//---------------------------------------------------------VFD
    // VTD (MOVI-C MOVIPRO) / Module 1 (Standard 8 PD), MOVIKIT Positioning Drive.
    // Raw 16-bit UINT data, as defined in SpaceX.tsproj; no scaling or decoding.
    // Link each variable to the channel with the same number in TwinCAT XAE.
    // Word meanings from MOVISUITE; bit meanings and units still pending SEW.

    // Drive -> PLC: Inputs 8 PD / PDO 16#1A02 / object 16#7002.
    // Read only by FC Inputs, into Control.VTD.Motor.stProcessInput.
    VTD_PI_01 AT %I* : UINT; // PI 1, 16#7002:01 - Status word
    VTD_PI_02 AT %I* : UINT; // PI 2, 16#7002:02 - Actual speed
    VTD_PI_03 AT %I* : UINT; // PI 3, 16#7002:03 - Status/main fault - subfault
    VTD_PI_04 AT %I* : UINT; // PI 4, 16#7002:04 - Torque
    VTD_PI_05 AT %I* : UINT; // PI 5, 16#7002:05 - Digital inputs
    VTD_PI_06 AT %I* : UINT; // PI 6, 16#7002:06 - Actual application mode
    VTD_PI_07 AT %I* : UINT; // PI 7, 16#7002:07 - Actual position high word (DL50)
    VTD_PI_08 AT %I* : UINT; // PI 8, 16#7002:08 - Actual position low word (DL50)

    // PLC -> drive: Outputs 8 PD / PDO 16#1602 / object 16#6002.
    // Written only by FC Outputs, from Control.VTD.Motor.aProcessOutput.
    VTD_PO_01 AT %Q* : UINT; // PO 1, 16#6002:01 - Control word
    VTD_PO_02 AT %Q* : UINT; // PO 2, 16#6002:02 - Setpoint speed
    VTD_PO_03 AT %Q* : UINT; // PO 3, 16#6002:03 - Setpoint acceleration
    VTD_PO_04 AT %Q* : UINT; // PO 4, 16#6002:04 - Setpoint deceleration
    VTD_PO_05 AT %Q* : UINT; // PO 5, 16#6002:05 - Digital outputs
    VTD_PO_06 AT %Q* : UINT; // PO 6, 16#6002:06 - Setpoint application mode
    VTD_PO_07 AT %Q* : UINT; // PO 7, 16#6002:07 - Target position high word
    VTD_PO_08 AT %Q* : UINT; // PO 8, 16#6002:08 - Target position low word

    // EtherCAT diagnostics of the VTD box. Not linked yet: link manually in XAE.
    // Read only by FC Inputs.
    VTD_WcState AT %I* : BOOL; // VTD > WcState > WcState (TRUE = data invalid)
    VTD_EcState AT %I* : UINT; // VTD > InfoData > State (8 = OP)
	
	//----------------------------------------------------EXTRACTOR CONVEYOR
END_VAR

// ---- GVLs/Settings.TcGVL
{attribute 'qualified_only'}
VAR_GLOBAL
	VTD:  VTD_Settings_DUT;
	ECnv:  ECnv_Settings_DUT;
	LCnv:  ARRAY[1..6] OF Buffer_Cnv_Settings_DUT;
	Turn_Table: Turn_Table_Settings_DUT;
	TBCnv:  TBCnv_Settings_DUT;
	Pop_Up_Cnv: ARRAY[1..2] OF PopUp_Settings_DUT;
	Roller_Cnv: ARRAY[1..5] OF Roller_Settings_DUT;
	Chain_Cnv: Chain_Settings_DUT;
// 	Shuttle_MQTT:  MQTT_Settings;
	System:  System_Settings_DUT;
END_VAR

// ---- GVLs/System.TcGVL
{attribute 'qualified_only'}
VAR_GLOBAL
	Id:  UINT;
	CancelOrders:  BOOL;
	PauseOrders:  Bool;
	ResumeOrders:  Bool;
	OrderSent:  Bool;
	CurrentOrder:  UInt;
	NextOrder:  UInt;
	OrderTable:  ARRAY[0..99] OF OrderTable_DUT;
	StepTable:  ARRAY[0..20] OF OrderTable_DUT;
	CarParked_Confirm:  Bool;
	Running:  Bool;
	IDLE:  Bool;
	Error:  Bool;
	State:  USInt;
	ResetError:  Bool;
	Ready:  Bool;
	Selected:  Bool;
	Auto_Man:  Bool;
	Paused:  Bool;
// 	Watchdog_TimeOut:  STRUCT;
END_VAR

// ---- GVLs/System_Control.TcGVL
{attribute 'qualified_only'}
VAR_GLOBAL
	Reset_All:  BOOL;
	MQTT_Enable:  BOOL;
	OPC_Enable:  Bool;
END_VAR

// ---- POUs/MAIN.TcPOU
PROGRAM MAIN
VAR
	 // TEST ONLY - VTD MOVIPRO process data communication check.
    fbVtdProcessDataTest : FB_SEW_ProcessDataTest;
    // TEST ONLY - VTD manual control from the screen VTD_ManualTest.
    fbVtdManualControl : FB_VTD_ManualControl;
    // Safety reset from the HMI (button SAFETY RESET): one pulse per rising edge.
    rtSafetyReset : R_TRIG;
    tpSafetyReset : TP;
END_VAR

run := TRUE;

// 1. IO inputs -> internal variables
Inputs();

// 2. Logic on internal variables
// Safety reset from the HMI: one 500 ms pulse on IO_Safety.ErrorAcknowledgement and
// IO_Safety.SEW_Safety_Reset (written in Outputs). It is a request only: the TwinSAFE
// logic accepts it or not. Holding the button does not repeat the reset.
rtSafetyReset(CLK := GVL_HMI_System.stCommand.bSafetyReset);
tpSafetyReset(IN := rtSafetyReset.Q, PT := T#500MS);
Control.SafetyReset := tpSafetyReset.Q;

// TEST ONLY - two sources can write the VTD process outputs, only one at a time:
//  - the raw write of the process data screen is refused (its HMI toggle is reset)
//    while the manual screen has the drive enabled;
//  - the manual control is inhibited while the raw write is active.
IF fbVtdManualControl.q_stStatus.bEnableActive THEN
    GVL_HMI_VTD.stPdCommand.bTestWriteEnable := FALSE;
END_IF

// TEST ONLY - VTD MOVIPRO process data communication check.
fbVtdProcessDataTest(
    i_aProcessInput := Control.VTD.Motor.stProcessInput.aWord,
    i_bWcStateError := Control.VTD.Motor.stProcessInput.bWcStateError,
    i_uiEcState := Control.VTD.Motor.stProcessInput.uiEcState,
    i_bTestWriteEnable := GVL_HMI_VTD.stPdCommand.bTestWriteEnable,
    i_bTestAllowControlWord := GVL_HMI_VTD.stPdCommand.bTestAllowControlWord,
    i_aTestProcessOutput := GVL_HMI_VTD.stPdCommand.aTestProcessOutput);

// TEST ONLY - VTD manual control (jog, modes, speed, software stop, reset).
fbVtdManualControl(
    i_stProcessInput := Control.VTD.Motor.stProcessInput,
    i_bInhibit := fbVtdProcessDataTest.q_bTestWriteActive,
    i_stSettings := GVL_HMI_VTD.stManualSettings,
    io_stCommand := GVL_HMI_VTD.stManualCommand);

IF fbVtdProcessDataTest.q_bTestWriteActive THEN
    Control.VTD.Motor.aProcessOutput := fbVtdProcessDataTest.q_aProcessOutput;
ELSE
    Control.VTD.Motor.aProcessOutput := fbVtdManualControl.q_aProcessOutput;
END_IF

// 3. HMI status
FC_VTD_PdHmiUpdateStatus(
    io_fbProcessData := fbVtdProcessDataTest,
    io_stStatus := GVL_HMI_VTD.stPdStatus);
// PO really sent to the drive (raw write or manual control).
GVL_HMI_VTD.stPdStatus.aProcessOutputSent := Control.VTD.Motor.aProcessOutput;
GVL_HMI_VTD.stManualStatus := fbVtdManualControl.q_stStatus;
GVL_HMI_System.stStatus.bSafetyResetActive := tpSafetyReset.Q;

// 4. Internal variables -> IO outputs
Outputs();

END_PROGRAM

// ---- POUs/SEW/FB_SEW_ProcessDataTest.TcPOU
// TEST ONLY - communication check between TwinCAT and a MOVIPRO running
// MOVIKIT Positioning Drive with the "Standard 8 PD" fieldbus interface.
//
// PD layout confirmed from MOVISUITE (VTD > MOVIKIT Positioning Drive > Basic settings):
//   PO 1 Control word              PI 1 Status word
//   PO 2 Setpoint speed            PI 2 Actual speed
//   PO 3 Setpoint acceleration     PI 3 Status/main fault - subfault
//   PO 4 Setpoint deceleration     PI 4 Torque (selectable in MOVISUITE)
//   PO 5 Digital outputs           PI 5 Digital inputs
//   PO 6 Setpoint application mode PI 6 Actual application mode
//   PO 7 Target position high word PI 7 Actual position high word
//   PO 8 Target position low word  PI 8 Actual position low word
//
// NOT yet confirmed (pending SEW): control/status word bit meanings,
// application mode values, user units and scaling of speed, ramps, torque and
// position. All decoded values are therefore RAW and carry no engineering unit.
//
// This block does not control the drive. All process outputs are 0 unless a
// TEST ONLY write is explicitly enabled online. The control word (PO 1) stays 0
// unless it is separately enabled. A control word of 0 is not confirmed as a
// safe state for this vertical axis; confirm with SEW before writing anything.
FUNCTION_BLOCK FB_SEW_ProcessDataTest
VAR_INPUT
    i_aProcessInput : ARRAY[1..8] OF UINT;      // PI 1..8, raw from the drive
    i_bWcStateError : BOOL;                     // EtherCAT WcState of the drive box (TRUE = data invalid)
    i_uiEcState : UINT;                         // EtherCAT InfoData.State of the drive box (8 = OP)

    i_bTestWriteEnable : BOOL;                  // TEST ONLY - allow PO 2..8 to be written
    i_bTestAllowControlWord : BOOL;             // TEST ONLY - additionally allow PO 1 (control word)
    i_aTestProcessOutput : ARRAY[1..8] OF UINT; // TEST ONLY - raw values to send to PO 1..8
    i_tTestWriteTimeout : TIME := T#10M;        // TEST ONLY write is dropped after this time
END_VAR
VAR_OUTPUT
    q_bCommunicationOk : BOOL;                  // Drive in OP and working counter valid
    q_udiInputChangeCount : UDINT;              // Cycles in which any PI word changed (wraps)

    q_wStatusWord : WORD;                       // PI 1, bit meanings pending SEW
    q_iActualSpeedRaw : INT;                    // PI 2, signed assumed, unit pending SEW
    q_wFaultCode : WORD;                        // PI 3, main fault / subfault, raw
    q_iTorqueRaw : INT;                         // PI 4, signed assumed, unit pending SEW
    q_wDigitalInputs : WORD;                    // PI 5, raw
    q_uiActualApplicationMode : UINT;           // PI 6, value meanings pending SEW
    q_diActualPositionRaw : DINT;               // PI 7 (high) + PI 8 (low), user units pending SEW

    q_bTestWriteActive : BOOL;                  // TEST ONLY write currently applied
    q_bTestWriteExpired : BOOL;                 // Timeout elapsed; toggle i_bTestWriteEnable to restart
    q_tTestWriteElapsed : TIME;                 // Elapsed time of the current TEST ONLY write window
    q_aProcessOutput : ARRAY[1..8] OF UINT;     // PO 1..8, raw to the drive
END_VAR
VAR
    aPreviousInput : ARRAY[1..8] OF UINT;
    bInputChanged : BOOL;
    dwActualPosition : DWORD;
    iWord : INT;

    rtrigTestWriteEnable : R_TRIG;
    tonTestWriteTimeout : TON;
END_VAR

// Communication status: EtherCAT state OP (lower nibble = 8) and valid working counter.
q_bCommunicationOk := (NOT i_bWcStateError) AND ((i_uiEcState AND 16#000F) = 8);

// Count cycles in which the drive sends new data. A counter that keeps rising
// while the drive is powered shows that PI data really arrives.
bInputChanged := FALSE;
FOR iWord := 1 TO 8 DO
    IF i_aProcessInput[iWord] <> aPreviousInput[iWord] THEN
        bInputChanged := TRUE;
    END_IF
END_FOR
aPreviousInput := i_aProcessInput;

IF bInputChanged THEN
    q_udiInputChangeCount := q_udiInputChangeCount + 1;
END_IF

// Raw decoding. Same-size integer conversions keep the bit pattern.
q_wStatusWord := UINT_TO_WORD(i_aProcessInput[1]);
q_iActualSpeedRaw := UINT_TO_INT(i_aProcessInput[2]);
q_wFaultCode := UINT_TO_WORD(i_aProcessInput[3]);
q_iTorqueRaw := UINT_TO_INT(i_aProcessInput[4]);
q_wDigitalInputs := UINT_TO_WORD(i_aProcessInput[5]);
q_uiActualApplicationMode := i_aProcessInput[6];

// Position word order (PI 7 = high, PI 8 = low) is shown in MOVISUITE.
// Signed 32-bit integer: numeric value, not an IEEE-754 bit pattern.
dwActualPosition := SHL(UINT_TO_DWORD(i_aProcessInput[7]), 16)
                    OR UINT_TO_DWORD(i_aProcessInput[8]);
q_diActualPositionRaw := DWORD_TO_DINT(dwActualPosition);

// TEST ONLY write enable with timeout. A rising edge restarts the timeout.
rtrigTestWriteEnable(CLK := i_bTestWriteEnable);
IF rtrigTestWriteEnable.Q THEN
    q_bTestWriteExpired := FALSE;
END_IF

tonTestWriteTimeout(IN := i_bTestWriteEnable AND NOT q_bTestWriteExpired,
                    PT := i_tTestWriteTimeout);
IF tonTestWriteTimeout.Q THEN
    q_bTestWriteExpired := TRUE;
END_IF
q_tTestWriteElapsed := tonTestWriteTimeout.ET;

q_bTestWriteActive := i_bTestWriteEnable AND NOT q_bTestWriteExpired;

// Process outputs: 0 by default.
FOR iWord := 1 TO 8 DO
    q_aProcessOutput[iWord] := 0;
END_FOR

IF q_bTestWriteActive THEN
    FOR iWord := 2 TO 8 DO
        q_aProcessOutput[iWord] := i_aTestProcessOutput[iWord];
    END_FOR

    IF i_bTestAllowControlWord THEN
        q_aProcessOutput[1] := i_aTestProcessOutput[1];
    END_IF
END_IF

END_FUNCTION_BLOCK

// ---- POUs/VTD/FB_VTD_ManualControl.TcPOU
// TEST ONLY - manual control of the VTD MOVIPRO from the screen VTD_ManualTest.
// Temporary owner of the axis for commissioning; VTD_FB replaces it in production.
// Uses FB_SEW_Drive (MOVIKIT Positioning Drive, Standard 8 PD, SEW manual 33959862).
//
// Behavior:
//  - ENABLE is a request from the HMI. It is dropped, and the HMI toggle reset, on
//    software stop, communication loss, drive error, STO active or while the raw
//    process data write is active. No automatic restart.
//    ENABLE off while turning: stop with the PO 4 ramp first, then remove the enable.
//  - JOG -/+ (modes 100/101) is hold-to-run. A button must be released before it is
//    accepted, and it is ignored after tJogMaxTime until it is released.
//  - RUN -/+ (mode 200) and START (modes 300/400/401) are latched; STOP clears them
//    (deceleration with PO 4). Reversing in mode 200 requires STOP first.
//  - The target position is taken from the HMI only with START.
//  - The operating mode changes only at standstill without motion command,
//    because the drive stops when PO 6 changes (manual chapter 8.1).
//  - Speed = iSpeedPercent (0..100 %) of stManualSettings.iMaxSpeed (user units).
//  - SOFTWARE STOP is NOT an emergency stop and not a safety function. It removes the
//    enable, so the drive stops with FCB 14 (emergency stop ramp) and applies the brake.
//    The safety-rated stop is the hardwired / TwinSAFE emergency stop (STO).
//  - RESET clears the software stop and sends a drive fault reset pulse (PO 1.8).
//  - Never used: release brake without enable, output stage inhibit, deactivation of
//    the software limit switches (not set by FB_SEW_Drive).
//
// Drive status is evaluated from the previous call of FB_SEW_Drive (one PLC cycle).
FUNCTION_BLOCK FB_VTD_ManualControl
VAR_INPUT
    i_stProcessInput : ST_SEW_ProcessInput8;  // Raw PI 1..8 + EtherCAT diagnostics (Control.VTD.Motor)
    i_bInhibit : BOOL;                        // TRUE = another source writes the PO (raw PD test); enable is dropped
    i_stSettings : ST_VTD_ManualSettings;     // Max speed, ramps (user units) and jog max time
END_VAR
VAR_IN_OUT
    io_stCommand : ST_VTD_ManualHmiCommand;   // HMI commands; bEnable, eModeRequest and iSpeedPercent are written back
END_VAR
VAR_OUTPUT
    q_aProcessOutput : ARRAY[1..8] OF UINT;   // Raw PO 1..8 (to Control.VTD.Motor.aProcessOutput)
    q_stStatus : ST_VTD_ManualHmiStatus;      // To GVL_HMI_VTD.stManualStatus
END_VAR
VAR
    fbDrive : FB_SEW_Drive;
    eModeActive : E_SEW_MovikitMode := E_SEW_MovikitMode.JogSpeedControlled;

    // Operating mode
    bModeSupported : BOOL;
    bModeChangeAllowed : BOOL;
    bModeRejected : BOOL;
    bJogMode : BOOL;
    bSpeedMode : BOOL;
    bReferencingMode : BOOL;
    bPositioningMode : BOOL;

    // Enable
    bSoftwareStopLatched : BOOL;
    bSettingsValid : BOOL;
    bEnableBlocked : BOOL;
    bEnableRequest : BOOL;
    bEnableActive : BOOL;

    // Motion commands
    bMotionCommand : BOOL;
    bJogButtonsReleased : BOOL;
    bJogArmed : BOOL;
    bJogTimeout : BOOL;
    bJogPositive : BOOL;
    bJogNegative : BOOL;
    bRunAvailable : BOOL;
    bRunPositive : BOOL;
    bRunNegative : BOOL;
    bStartAvailable : BOOL;
    bStartLatched : BOOL;
    bRelativeMoveOpen : BOOL;                 // Mode 401: distance applied, target not reached yet
    bApplyRelativeRequest : BOOL;             // Mode 401: PO 1.6 pulse starts in the next cycle
    diTargetPosition : DINT;                  // PO 7/8, user units
    diSpeedTemp : DINT;
    iSpeedMagnitude : INT;
    iSpeedSetpoint : INT;

    rtrigSoftwareStop : R_TRIG;
    rtrigReset : R_TRIG;
    rtrigRunPositive : R_TRIG;
    rtrigRunNegative : R_TRIG;
    rtrigStart : R_TRIG;
    rtrigStop : R_TRIG;
    tpFaultReset : TP;
    tpApplyRelative : TP;
    tpModeRejected : TP;
    tonJogMaxTime : TON;
    tonDisableStop : TON;
    tonRelativeDone : TON;
    tonReferencingDone : TON;
END_VAR
VAR CONSTANT
    FAULT_RESET_PULSE : TIME := T#500MS;      // PO 1.8 high time (the drive resets on the rising edge)
    APPLY_RELATIVE_PULSE : TIME := T#200MS;   // PO 1.6 high time (mode 401)
    MODE_REJECTED_MESSAGE : TIME := T#3S;     // Display time of the "mode change refused" message
    DISABLE_STOP_TIMEOUT : TIME := T#5S;      // Max time to stop with PO 4 before the enable is removed
    RELATIVE_DONE_DELAY : TIME := T#500MS;    // In position + standstill for this time = relative move done
    REFERENCING_DONE_DELAY : TIME := T#1S;    // Referenced + standstill for this time = START released
END_VAR

{region "Edge detection of the HMI buttons"}
rtrigSoftwareStop(CLK := io_stCommand.bSoftwareStop);
rtrigReset(CLK := io_stCommand.bReset);
rtrigRunPositive(CLK := io_stCommand.bRunPositive);
rtrigRunNegative(CLK := io_stCommand.bRunNegative);
rtrigStart(CLK := io_stCommand.bStart);
rtrigStop(CLK := io_stCommand.bStop);
{endregion}

{region "Software stop and reset"}
// SOFTWARE STOP is not a safety function. It removes the enable, so the drive
// stops with FCB 14 (emergency stop ramp) and applies the brake.
IF rtrigSoftwareStop.Q THEN
    bSoftwareStopLatched := TRUE;
END_IF

// RESET clears the software stop and resets drive faults with a PO 1.8 pulse.
// The enable stays off until ENABLE is pressed again.
IF rtrigReset.Q AND NOT io_stCommand.bSoftwareStop THEN
    bSoftwareStopLatched := FALSE;
END_IF
tpFaultReset(IN := rtrigReset.Q, PT := FAULT_RESET_PULSE);
{endregion}

{region "Settings"}
bSettingsValid := (i_stSettings.iMaxSpeed > 0)
                  AND (i_stSettings.uiAcceleration > 0)
                  AND (i_stSettings.uiDeceleration > 0)
                  AND (i_stSettings.tJogMaxTime > T#0S);
{endregion}

{region "Operating mode (PO 6)"}
// The drive stops when PO 6 changes (manual chapter 8.1), so the mode is changed
// only at standstill and without an active motion command.
bMotionCommand := bRunPositive OR bRunNegative OR bStartLatched
                  OR io_stCommand.bJogPositive OR io_stCommand.bJogNegative;
bModeChangeAllowed := NOT bMotionCommand AND NOT fbDrive.q_stStatus.bMotorTurning;
bModeRejected := FALSE;

IF io_stCommand.eModeRequest <> eModeActive THEN
    CASE io_stCommand.eModeRequest OF
        E_SEW_MovikitMode.JogPositionControlled,
        E_SEW_MovikitMode.JogSpeedControlled,
        E_SEW_MovikitMode.Speed,
        E_SEW_MovikitMode.ReferencingOffsetConfigured,
        E_SEW_MovikitMode.PositioningAbsolute,
        E_SEW_MovikitMode.PositioningRelative:
            bModeSupported := TRUE;
    ELSE
        bModeSupported := FALSE;
    END_CASE

    IF bModeSupported AND bModeChangeAllowed THEN
        eModeActive := io_stCommand.eModeRequest;
        bRelativeMoveOpen := FALSE;
        diTargetPosition := 0;
    ELSE
        bModeRejected := TRUE;
    END_IF
END_IF

// The HMI always shows the mode really sent to the drive.
io_stCommand.eModeRequest := eModeActive;

bJogMode := (eModeActive = E_SEW_MovikitMode.JogPositionControlled)
            OR (eModeActive = E_SEW_MovikitMode.JogSpeedControlled);
bSpeedMode := (eModeActive = E_SEW_MovikitMode.Speed);
bReferencingMode := (eModeActive = E_SEW_MovikitMode.ReferencingOffsetConfigured);
bPositioningMode := (eModeActive = E_SEW_MovikitMode.PositioningAbsolute)
                    OR (eModeActive = E_SEW_MovikitMode.PositioningRelative);
{endregion}

{region "Enable (PO 1.0 + PO 1.1)"}
// The enable request is dropped - and the HMI toggle reset - when the drive cannot
// or must not run. No automatic restart: ENABLE must be pressed again.
bEnableBlocked := bSoftwareStopLatched
                  OR i_bInhibit
                  OR NOT fbDrive.q_stStatus.bCommunicationOk
                  OR fbDrive.q_stStatus.bError
                  OR NOT fbDrive.q_stStatus.bStoInactive;

IF bEnableBlocked THEN
    io_stCommand.bEnable := FALSE;
END_IF
bEnableRequest := io_stCommand.bEnable AND NOT bEnableBlocked;

// ENABLE switched off while turning: the motion commands are cleared below, the
// drive stops with the PO 4 ramp and the enable is removed at standstill
// (at the latest after DISABLE_STOP_TIMEOUT, then FCB 14).
tonDisableStop(IN := bEnableActive AND NOT bEnableRequest AND NOT bEnableBlocked,
               PT := DISABLE_STOP_TIMEOUT);
bEnableActive := bEnableRequest
                 OR (bEnableActive
                     AND NOT bEnableBlocked
                     AND fbDrive.q_stStatus.bMotorTurning
                     AND NOT tonDisableStop.Q);

// Manual chapter 8.1.8: after the enable was removed, a relative move must be
// started again with "Apply relative position".
IF NOT bEnableActive THEN
    bRelativeMoveOpen := FALSE;
END_IF
{endregion}

{region "JOG -/+ (modes 100/101) - hold-to-run"}
bJogButtonsReleased := NOT io_stCommand.bJogPositive AND NOT io_stCommand.bJogNegative;

// A jog button is accepted only after both buttons were released while jog was
// possible, so a button held during ENABLE or a mode change does not move the axis.
IF NOT (bEnableRequest AND bJogMode AND bSettingsValid) THEN
    bJogArmed := FALSE;
ELSIF bJogButtonsReleased THEN
    bJogArmed := TRUE;
END_IF

// Max continuous jog time. Also limits a jog left active by a lost HMI connection.
tonJogMaxTime(IN := NOT bJogButtonsReleased, PT := i_stSettings.tJogMaxTime);
IF tonJogMaxTime.Q THEN
    bJogTimeout := TRUE;
ELSIF bJogButtonsReleased THEN
    bJogTimeout := FALSE;
END_IF

bJogPositive := bJogArmed AND NOT bJogTimeout
                AND io_stCommand.bJogPositive AND NOT io_stCommand.bJogNegative;
bJogNegative := bJogArmed AND NOT bJogTimeout
                AND io_stCommand.bJogNegative AND NOT io_stCommand.bJogPositive;
{endregion}

{region "RUN -/+ (mode 200) - latched"}
bRunAvailable := bEnableRequest AND bSpeedMode AND bSettingsValid;

IF NOT bRunAvailable OR rtrigStop.Q THEN
    bRunPositive := FALSE;
    bRunNegative := FALSE;
ELSIF rtrigRunPositive.Q AND NOT bRunNegative THEN
    bRunPositive := TRUE;
ELSIF rtrigRunNegative.Q AND NOT bRunPositive THEN
    bRunNegative := TRUE;
END_IF
{endregion}

{region "START (modes 300/400/401) - latched"}
// PO 1.6 pulse for mode 401, requested in the previous cycle (PO 7/8 already sent).
tpApplyRelative(IN := bApplyRelativeRequest, PT := APPLY_RELATIVE_PULSE);
bApplyRelativeRequest := FALSE;

bStartAvailable := bEnableRequest AND bSettingsValid
                   AND (bReferencingMode
                        OR (bPositioningMode AND fbDrive.q_stStatus.bReferenced));

IF NOT bStartAvailable OR rtrigStop.Q THEN
    bStartLatched := FALSE;
ELSIF rtrigStart.Q THEN
    IF eModeActive = E_SEW_MovikitMode.PositioningRelative THEN
        IF bRelativeMoveOpen THEN
            // Move interrupted with STOP: continue to the original target (manual 8.1.8).
            bStartLatched := TRUE;
        ELSIF NOT fbDrive.q_stStatus.bMotorTurning THEN
            // New relative move: distance in PO 7/8 now, PO 1.6 edge from the next cycle.
            diTargetPosition := io_stCommand.diTargetPosition;
            bApplyRelativeRequest := TRUE;
            bRelativeMoveOpen := TRUE;
            bStartLatched := TRUE;
        END_IF
    ELSIF eModeActive = E_SEW_MovikitMode.PositioningAbsolute THEN
        // Absolute target, taken from the HMI only now (PO 7/8 is applied live by the drive).
        diTargetPosition := io_stCommand.diTargetPosition;
        bStartLatched := TRUE;
    ELSE
        // Referencing (300): offset from the MOVISUITE configuration, PO 7/8 not used.
        bStartLatched := TRUE;
    END_IF
END_IF

// Relative move finished: in position and standstill for RELATIVE_DONE_DELAY.
tonRelativeDone(IN := bRelativeMoveOpen AND bStartLatched AND NOT tpApplyRelative.Q
                      AND fbDrive.q_stStatus.bInPosition
                      AND NOT fbDrive.q_stStatus.bMotorTurning,
                PT := RELATIVE_DONE_DELAY);
IF tonRelativeDone.Q THEN
    bRelativeMoveOpen := FALSE;
END_IF

// Referencing finished: referenced and standstill -> START is released.
tonReferencingDone(IN := bStartLatched AND bReferencingMode
                         AND fbDrive.q_stStatus.bReferenced
                         AND NOT fbDrive.q_stStatus.bMotorTurning,
                   PT := REFERENCING_DONE_DELAY);
IF tonReferencingDone.Q THEN
    bStartLatched := FALSE;
END_IF
{endregion}

{region "Speed setpoint (PO 2)"}
io_stCommand.iSpeedPercent := LIMIT(0, io_stCommand.iSpeedPercent, 100);

diSpeedTemp := INT_TO_DINT(i_stSettings.iMaxSpeed) * INT_TO_DINT(io_stCommand.iSpeedPercent) / 100;
iSpeedMagnitude := DINT_TO_INT(LIMIT(0, diSpeedTemp, 32767));

// Signed only in mode 200 (RUN -); jog and positioning use the magnitude.
IF bRunNegative THEN
    iSpeedSetpoint := -iSpeedMagnitude;
ELSE
    iSpeedSetpoint := iSpeedMagnitude;
END_IF
{endregion}

{region "SEW communication layer"}
fbDrive(
    i_stProcessInput := i_stProcessInput,
    i_bEnable := bEnableActive,
    i_bStart := bRunPositive OR bRunNegative OR bStartLatched,
    i_bJogPositive := bJogPositive,
    i_bJogNegative := bJogNegative,
    i_bApplyRelativePosition := tpApplyRelative.Q,
    i_bFaultReset := tpFaultReset.Q,
    i_eMode := eModeActive,
    i_iSpeedSetpoint := iSpeedSetpoint,
    i_uiAcceleration := i_stSettings.uiAcceleration,
    i_uiDeceleration := i_stSettings.uiDeceleration,
    i_diTargetPosition := diTargetPosition);

q_aProcessOutput := fbDrive.q_aProcessOutput;
{endregion}

{region "HMI status"}
tpModeRejected(IN := bModeRejected, PT := MODE_REJECTED_MESSAGE);

q_stStatus.stDrive := fbDrive.q_stStatus;
q_stStatus.udiErrorId := fbDrive.q_udiErrorId;
q_stStatus.sActualModeName := FC_SEW_MovikitModeName(i_uiMode := fbDrive.q_stStatus.uiActualMode);

q_stStatus.eModeActive := eModeActive;
q_stStatus.sModeActiveName := FC_SEW_MovikitModeName(i_uiMode := TO_UINT(eModeActive));
q_stStatus.bModeJogPosition := (eModeActive = E_SEW_MovikitMode.JogPositionControlled);
q_stStatus.bModeJogSpeed := (eModeActive = E_SEW_MovikitMode.JogSpeedControlled);
q_stStatus.bModeSpeed := bSpeedMode;
q_stStatus.bModeReferencing := bReferencingMode;
q_stStatus.bModePositionAbsolute := (eModeActive = E_SEW_MovikitMode.PositioningAbsolute);
q_stStatus.bModePositionRelative := (eModeActive = E_SEW_MovikitMode.PositioningRelative);
q_stStatus.bModeChangeAllowed := bModeChangeAllowed;

q_stStatus.bEnableActive := bEnableActive;
q_stStatus.bSoftwareStopActive := bSoftwareStopLatched;
q_stStatus.bRawWriteActive := i_bInhibit;
q_stStatus.bSettingsValid := bSettingsValid;
q_stStatus.bJogAvailable := bEnableRequest AND bJogMode AND bSettingsValid;
q_stStatus.bRunAvailable := bRunAvailable;
q_stStatus.bStartAvailable := bStartAvailable;
q_stStatus.bJogPositiveActive := bJogPositive;
q_stStatus.bJogNegativeActive := bJogNegative;
q_stStatus.bJogTimeout := bJogTimeout;
q_stStatus.bRunPositiveActive := bRunPositive;
q_stStatus.bRunNegativeActive := bRunNegative;
q_stStatus.bStartActive := bStartLatched;
q_stStatus.bFaultResetActive := tpFaultReset.Q;

q_stStatus.iSpeedSetpoint := UINT_TO_INT(q_aProcessOutput[2]);
q_stStatus.diTargetPositionSent := diTargetPosition;

// Operator message: stop/fault conditions first (red), then hints.
q_stStatus.bMessageAlarm := TRUE;
IF i_bInhibit THEN
    q_stStatus.sMessage := 'Raw PD write active on the process data screen - switch it off';
ELSIF NOT fbDrive.q_stStatus.bCommunicationOk THEN
    q_stStatus.sMessage := 'No communication with the drive (EtherCAT or MOVIKIT handshake)';
ELSIF bSoftwareStopLatched THEN
    q_stStatus.sMessage := 'SOFTWARE STOP active - press RESET';
ELSIF NOT fbDrive.q_stStatus.bStoInactive THEN
    q_stStatus.sMessage := 'STO active - check emergency stop / safety circuit';
ELSIF fbDrive.q_stStatus.bError THEN
    q_stStatus.sMessage := 'Drive fault - see fault code, press RESET';
ELSIF NOT bSettingsValid THEN
    q_stStatus.sMessage := 'Enter max speed, acceleration and deceleration (test settings)';
ELSE
    q_stStatus.bMessageAlarm := FALSE;
    IF tpModeRejected.Q THEN
        q_stStatus.sMessage := 'Mode change refused - press STOP and wait for standstill';
    ELSIF bJogTimeout THEN
        q_stStatus.sMessage := 'Jog time limit reached - release the jog button';
    ELSIF bPositioningMode AND NOT fbDrive.q_stStatus.bReferenced THEN
        q_stStatus.sMessage := 'Axis not referenced - use mode 300 first';
    ELSIF NOT bEnableActive THEN
        q_stStatus.sMessage := 'Press ENABLE';
    ELSE
        q_stStatus.sMessage := 'Ready';
    END_IF
END_IF
{endregion}

END_FUNCTION_BLOCK

// ---- POUs/SEW/FB_SEW_Drive.TcPOU
// Communication and status layer for a SEW drive running MOVIKIT Positioning
// with the "Standard 8 PD" fieldbus interface (SBusPLUS, not CiA402).
// Source: SEW manual 33959862, chapter 9 "Process data assignment".
//
// This block does NOT decide any motion. The owner of the axis (e.g. VTD_FB)
// sets the commands; this block only packs them into PO 1..8, decodes PI 1..8
// and supervises the communication (EtherCAT state + MOVIKIT handshake).
//
// Safety-related behavior:
//  - Enable, start and jog are forced to 0 while communication is not OK.
//  - PO 1.3 "Release brake (without enable)" is never set (vertical axis).
//  - PO 1.13 "Output stage inhibit" is never set; removing enable stops the
//    drive with the emergency stop ramp (FCB 14) and applies the brake.
FUNCTION_BLOCK FB_SEW_Drive
VAR_INPUT
    i_stProcessInput : ST_SEW_ProcessInput8;  // Raw PI 1..8 + EtherCAT diagnostics (from FC Inputs)

    i_bEnable : BOOL;                         // PO 1.0 + PO 1.1 enable (FALSE = stop with FCB 14)
    i_bStart : BOOL;                          // PO 1.7 start/stop with fieldbus ramp
    i_bJogPositive : BOOL;                    // PO 1.4, jog modes only
    i_bJogNegative : BOOL;                    // PO 1.5, jog modes only
    i_bApplyRelativePosition : BOOL;          // PO 1.6, mode 401 only, the drive applies PO 7/8 on the rising edge
    i_bFaultReset : BOOL;                     // PO 1.8, drive resets on the rising edge
    i_eMode : E_SEW_MovikitMode;              // PO 6 setpoint application mode

    i_iSpeedSetpoint : INT;                   // PO 2, signed, user units
    i_uiAcceleration : UINT;                  // PO 3, user units
    i_uiDeceleration : UINT;                  // PO 4, user units
    i_diTargetPosition : DINT;                // PO 7 (high) + PO 8 (low), user units

    i_tHandshakeTimeout : TIME := T#1S;       // Max time for PI 1.15 to follow PO 1.15
END_VAR
VAR_OUTPUT
    q_aProcessOutput : ARRAY[1..8] OF UINT;   // Raw PO 1..8 (to FC Outputs)
    q_stStatus : ST_SEW_MovikitStatus;        // Decoded PI 1..8

    q_bReady : BOOL;                          // Communication OK, ready, STO inactive, no error
    q_bError : BOOL;                          // Drive error or communication error
    q_udiErrorId : UDINT;                     // See ERROR_ID_* below, or PI 3 (fault * 256 + subfault)
END_VAR
VAR
    bHandshakeIn : BOOL;                      // Value sent in PO 1.15
    bHandshakeWaiting : BOOL;
    tonHandshake : TON;
    wControlWord : WORD;
    dwTargetPosition : DWORD;
    dwActualPosition : DWORD;
END_VAR
VAR CONSTANT
    ERROR_ID_ETHERCAT : UDINT := 16#FFFF0001; // Drive not in OP or working counter invalid
    ERROR_ID_HANDSHAKE : UDINT := 16#FFFF0002; // MOVIKIT handshake timeout
END_VAR

{region "Communication supervision"}
// EtherCAT: state OP (lower nibble = 8) and valid working counter.
q_stStatus.bEtherCatOk := (NOT i_stProcessInput.bWcStateError)
                          AND ((i_stProcessInput.uiEcState AND 16#000F) = 8);

// MOVIKIT handshake (manual chapter 9.3): the drive copies PO 1.15 to PI 1.15.
// When both are equal, invert PO 1.15; otherwise the timeout runs.
q_stStatus.bHandshakeOut := i_stProcessInput.aWord[1].15;

IF q_stStatus.bEtherCatOk THEN
    IF bHandshakeIn = q_stStatus.bHandshakeOut THEN
        bHandshakeIn := NOT bHandshakeIn;
        bHandshakeWaiting := FALSE;
    ELSE
        bHandshakeWaiting := TRUE;
    END_IF
ELSE
    // No valid data: the EtherCAT error is reported instead of the handshake.
    bHandshakeWaiting := FALSE;
END_IF

tonHandshake(IN := bHandshakeWaiting, PT := i_tHandshakeTimeout);
q_stStatus.bHandshakeError := tonHandshake.Q;

q_stStatus.bCommunicationOk := q_stStatus.bEtherCatOk AND NOT q_stStatus.bHandshakeError;
{endregion}

{region "Decode process inputs (PI 1..8)"}
q_stStatus.wStatusWord := UINT_TO_WORD(i_stProcessInput.aWord[1]);
q_stStatus.bReady := q_stStatus.wStatusWord.0;
q_stStatus.bStoInactive := q_stStatus.wStatusWord.1;
q_stStatus.bOutputStageEnabled := q_stStatus.wStatusWord.2;
q_stStatus.bBrakeReleased := q_stStatus.wStatusWord.3;
q_stStatus.bMotorTurning := q_stStatus.wStatusWord.4;
q_stStatus.bReferenced := q_stStatus.wStatusWord.5;
q_stStatus.bRelativePositionApplied := q_stStatus.wStatusWord.6;
q_stStatus.bInPosition := q_stStatus.wStatusWord.7;
q_stStatus.bError := q_stStatus.wStatusWord.8;
q_stStatus.bWarning := q_stStatus.wStatusWord.9;
q_stStatus.bDriveTrain2Active := q_stStatus.wStatusWord.10;
q_stStatus.bSpeedReached := q_stStatus.wStatusWord.11;
q_stStatus.bSwLimitSwitchesInactive := q_stStatus.wStatusWord.12;
q_stStatus.bStandbyActive := q_stStatus.wStatusWord.14;

// Same-size integer conversions keep the bit pattern (signed values).
q_stStatus.iActualSpeed := UINT_TO_INT(i_stProcessInput.aWord[2]);
q_stStatus.byFaultCode := WORD_TO_BYTE(SHR(UINT_TO_WORD(i_stProcessInput.aWord[3]), 8));
q_stStatus.bySubfaultCode := WORD_TO_BYTE(UINT_TO_WORD(i_stProcessInput.aWord[3]) AND 16#00FF);
q_stStatus.iActualTorque_0p1pct := UINT_TO_INT(i_stProcessInput.aWord[4]);
q_stStatus.wDigitalInputs := UINT_TO_WORD(i_stProcessInput.aWord[5]);
q_stStatus.uiActualMode := i_stProcessInput.aWord[6];

// Position: PI 7 = high word, PI 8 = low word, signed 32-bit integer (numeric, not REAL).
dwActualPosition := SHL(UINT_TO_DWORD(i_stProcessInput.aWord[7]), 16)
                    OR UINT_TO_DWORD(i_stProcessInput.aWord[8]);
q_stStatus.diActualPosition := DWORD_TO_DINT(dwActualPosition);
{endregion}

{region "Diagnostics"}
q_bError := q_stStatus.bError OR NOT q_stStatus.bCommunicationOk;
q_bReady := q_stStatus.bCommunicationOk AND q_stStatus.bReady
            AND q_stStatus.bStoInactive AND NOT q_stStatus.bError;

IF NOT q_stStatus.bEtherCatOk THEN
    q_udiErrorId := ERROR_ID_ETHERCAT;
ELSIF q_stStatus.bHandshakeError THEN
    q_udiErrorId := ERROR_ID_HANDSHAKE;
ELSIF q_stStatus.bError THEN
    q_udiErrorId := UINT_TO_UDINT(i_stProcessInput.aWord[3]);
ELSE
    q_udiErrorId := 0;
END_IF
{endregion}

{region "Build process outputs (PO 1..8)"}
wControlWord := 0;

IF q_stStatus.bCommunicationOk AND i_bEnable THEN
    wControlWord.0 := TRUE;     // Enable/emergency stop
    wControlWord.1 := TRUE;     // Enable/application stop
    wControlWord.4 := i_bJogPositive AND NOT i_bJogNegative;
    wControlWord.5 := i_bJogNegative AND NOT i_bJogPositive;
    wControlWord.6 := i_bApplyRelativePosition; // Ineffective in modes other than 401
    wControlWord.7 := i_bStart; // Start/stop with fieldbus ramp
END_IF

wControlWord.8 := i_bFaultReset;  // Allowed without enable
wControlWord.15 := bHandshakeIn;  // MOVIKIT handshake, no effect on motion
// Never set: bit 3 (release brake without enable), bit 13 (output stage inhibit),
// bit 12 (deactivate SW limit switches), bit 10 (drive train 2), bit 14 (standby).

q_aProcessOutput[1] := WORD_TO_UINT(wControlWord);

IF q_stStatus.bCommunicationOk AND i_bEnable THEN
    q_aProcessOutput[2] := INT_TO_UINT(i_iSpeedSetpoint);
ELSE
    q_aProcessOutput[2] := 0;
END_IF

q_aProcessOutput[3] := i_uiAcceleration;
q_aProcessOutput[4] := i_uiDeceleration;
q_aProcessOutput[5] := 0;  // Drive digital outputs not used
q_aProcessOutput[6] := TO_UINT(i_eMode);

dwTargetPosition := DINT_TO_DWORD(i_diTargetPosition);
q_aProcessOutput[7] := DWORD_TO_UINT(SHR(dwTargetPosition, 16));
q_aProcessOutput[8] := DWORD_TO_UINT(dwTargetPosition AND 16#0000FFFF);
{endregion}

END_FUNCTION_BLOCK

// ---- POUs/Inputs.TcPOU
// Input mapping: the only place where PLC IO inputs are read.
// Copies IO GVL variables to internal variables (GVL Control). One region per device.
// Called first in MAIN.
FUNCTION Inputs : BOOL
VAR_INPUT
END_VAR
VAR
END_VAR

{region "Chargers - PROFINET (EL6633)"}
// TODO: unfinished, kept disabled so the project builds. Before enabling:
//  - confirm the charger byte order and REAL representation (DWORD_REAL body is commented out)
//  - Control.Charger_Level is ARRAY[2..6]; index [1] is out of range
//  - IO_Chargers.Inputs_1 is not linked in SpaceX.tsproj
// Original line, unchanged:
// Control.Charger_Level[1].Output_Voltage :=  DWORD_REAL(b0:= IO_Chargers.Inputs_1[0],b1:=IO_Chargers.Inputs_1[1],b2:=IO_Chargers.Inputs_1[2],b3:=IO_Chargers.Inputs_1[3],
{endregion}

{region "VTD 1 - MOVIPRO process inputs (SEW Standard 8 PD)"}
Control.VTD.Motor.stProcessInput.aWord[1] := IO_VFDs.VTD_PI_01; // Status word
Control.VTD.Motor.stProcessInput.aWord[2] := IO_VFDs.VTD_PI_02; // Actual speed
Control.VTD.Motor.stProcessInput.aWord[3] := IO_VFDs.VTD_PI_03; // Status/main fault - subfault
Control.VTD.Motor.stProcessInput.aWord[4] := IO_VFDs.VTD_PI_04; // Torque
Control.VTD.Motor.stProcessInput.aWord[5] := IO_VFDs.VTD_PI_05; // Digital inputs
Control.VTD.Motor.stProcessInput.aWord[6] := IO_VFDs.VTD_PI_06; // Actual application mode
Control.VTD.Motor.stProcessInput.aWord[7] := IO_VFDs.VTD_PI_07; // Actual position high word
Control.VTD.Motor.stProcessInput.aWord[8] := IO_VFDs.VTD_PI_08; // Actual position low word

Control.VTD.Motor.stProcessInput.bWcStateError := IO_VFDs.VTD_WcState;
Control.VTD.Motor.stProcessInput.uiEcState := IO_VFDs.VTD_EcState;
{endregion}

Inputs := TRUE;

END_FUNCTION

// ---- POUs/Outputs.TcPOU
// Output mapping: the only place where PLC IO outputs are written.
// Copies internal variables (GVL Control) to IO GVL variables. One region per device.
// Called last in MAIN.
FUNCTION Outputs : BOOL
VAR_INPUT
END_VAR
VAR
END_VAR

{region "VTD 1 - MOVIPRO process outputs (SEW Standard 8 PD)"}
IO_VFDs.VTD_PO_01 := Control.VTD.Motor.aProcessOutput[1]; // Control word
IO_VFDs.VTD_PO_02 := Control.VTD.Motor.aProcessOutput[2]; // Setpoint speed
IO_VFDs.VTD_PO_03 := Control.VTD.Motor.aProcessOutput[3]; // Setpoint acceleration
IO_VFDs.VTD_PO_04 := Control.VTD.Motor.aProcessOutput[4]; // Setpoint deceleration
IO_VFDs.VTD_PO_05 := Control.VTD.Motor.aProcessOutput[5]; // Digital outputs
IO_VFDs.VTD_PO_06 := Control.VTD.Motor.aProcessOutput[6]; // Setpoint application mode
IO_VFDs.VTD_PO_07 := Control.VTD.Motor.aProcessOutput[7]; // Target position high word
IO_VFDs.VTD_PO_08 := Control.VTD.Motor.aProcessOutput[8]; // Target position low word
{endregion}

{region "Safety - reset request to the TwinSAFE logic (standard PLC -> safety)"}
IO_Safety.ErrorAcknowledgement := Control.SafetyReset; // TwinSAFE group ErrAck
IO_Safety.SEW_Safety_Reset := Control.SafetyReset;     // TwinSAFE alias Safety_SEW_Reset
{endregion}

Outputs := TRUE;

END_FUNCTION

// ---- POUs/SEW/FC_SEW_MovikitModeName.TcPOU
// Readable name of a MOVIKIT operating mode value (PI 6 / PO 6), for HMI and diagnostics.
FUNCTION FC_SEW_MovikitModeName : STRING(40)
VAR_INPUT
    i_uiMode : UINT;
END_VAR

CASE i_uiMode OF
    0:   FC_SEW_MovikitModeName := 'Default (0)';
    100: FC_SEW_MovikitModeName := 'Jog position-controlled (100)';
    101: FC_SEW_MovikitModeName := 'Jog speed-controlled (101)';
    200: FC_SEW_MovikitModeName := 'Speed (200)';
    300: FC_SEW_MovikitModeName := 'Referencing offset configured (300)';
    301: FC_SEW_MovikitModeName := 'Referencing offset fieldbus (301)';
    400: FC_SEW_MovikitModeName := 'Positioning absolute (400)';
    401: FC_SEW_MovikitModeName := 'Positioning relative (401)';
    402: FC_SEW_MovikitModeName := 'Positioning modulo positive (402)';
    403: FC_SEW_MovikitModeName := 'Positioning modulo negative (403)';
    404: FC_SEW_MovikitModeName := 'Positioning modulo short (404)';
    420: FC_SEW_MovikitModeName := 'Touchprobe absolute direction (420)';
    421: FC_SEW_MovikitModeName := 'Touchprobe absolute sign (421)';
    422: FC_SEW_MovikitModeName := 'Touchprobe endless direction (422)';
    423: FC_SEW_MovikitModeName := 'Touchprobe endless sign (423)';
    700: FC_SEW_MovikitModeName := 'Brake test (700)';
ELSE
    FC_SEW_MovikitModeName := CONCAT('Unknown (', CONCAT(UINT_TO_STRING(i_uiMode), ')'));
END_CASE

END_FUNCTION

// ---- POUs/SEW/FC_VTD_PdHmiUpdateStatus.TcPOU
// HMI layer: copies the process data test results to the HMI status structure.
// Read only towards the FB; it never changes FB inputs or drive outputs.
FUNCTION FC_VTD_PdHmiUpdateStatus : BOOL
VAR_IN_OUT
    io_fbProcessData : FB_SEW_ProcessDataTest;
    io_stStatus : ST_VTD_PdHmiStatus;
END_VAR

// Communication
io_stStatus.bCommunicationOk := io_fbProcessData.q_bCommunicationOk;
io_stStatus.bWcStateError := io_fbProcessData.i_bWcStateError;
io_stStatus.uiEcState := io_fbProcessData.i_uiEcState;
io_stStatus.udiInputChangeCount := io_fbProcessData.q_udiInputChangeCount;

// Process inputs
io_stStatus.aProcessInputRaw := io_fbProcessData.i_aProcessInput;
io_stStatus.wStatusWord := io_fbProcessData.q_wStatusWord;
io_stStatus.iActualSpeedRaw := io_fbProcessData.q_iActualSpeedRaw;
io_stStatus.wFaultCode := io_fbProcessData.q_wFaultCode;
io_stStatus.iTorqueRaw := io_fbProcessData.q_iTorqueRaw;
io_stStatus.wDigitalInputs := io_fbProcessData.q_wDigitalInputs;
io_stStatus.uiActualApplicationMode := io_fbProcessData.q_uiActualApplicationMode;
io_stStatus.sActualModeName := FC_SEW_MovikitModeName(i_uiMode := io_fbProcessData.q_uiActualApplicationMode);
io_stStatus.diActualPositionRaw := io_fbProcessData.q_diActualPositionRaw;

// TEST ONLY write
io_stStatus.bTestWriteActive := io_fbProcessData.q_bTestWriteActive;
io_stStatus.bTestWriteExpired := io_fbProcessData.q_bTestWriteExpired;
io_stStatus.tTestWriteElapsed := io_fbProcessData.q_tTestWriteElapsed;
io_stStatus.aProcessOutputSent := io_fbProcessData.q_aProcessOutput;

FC_VTD_PdHmiUpdateStatus := TRUE;

END_FUNCTION

// ---- POUs/Conveyors/Buffer_Conveyor_FB.TcPOU
FUNCTION_BLOCK Buffer_Conveyor_FB
VAR_INPUT
	Cnv_Settings:  Buffer_Cnv_Settings_DUT;
	VTD_Level:  UINT;
	Safety_OK:  Bool;
	CNV_In_Out:  Bool;
	CNV1_2_Selected:  UInt;
	Time_CheckPallet:  Time;
	Time_CheckNoPallet:  TIME;
END_VAR
VAR_OUTPUT
END_VAR
VAR_IN_OUT
	Cnv_Control:  Buffer_Cnv_Control_DUT;
END_VAR
VAR
	State:  UINT;
	Timer_Transfer:  TON;
	Watchdog:  TON;
	Transfer_Direction:  String;
	MainSetpoint:  Int;
	R_Automatic_Mode:  R_TRIG;
	R_Start_DB:  R_TRIG;
	R_Stop_DB:  R_TRIG;
	ID_Decoded:  ID_Decoded_DUT;
	ID_Decoded_From:  ID_Decoded_DUT;
	ID_Decoded_To:  ID_Decoded_DUT;
	T_Ramp:  TON;
	HMI_Reset:  Bool;
	T_CheckNoPallet:  TON;
	Time_SlowDown_Ramp:  Time;
	T_CheckPallet:  TON;

	// SEW MOVIKIT Velocity Drive (region "VFD")
	fbVelocityDrive:  FB_SEW_VelocityDrive;
	bDriveMoveRequest:  BOOL;
	bDriveEnable:  BOOL;
	bDriveFaultReset:  BOOL;
	bDriveParamsValid:  BOOL;             // SEW scaling and ramps configured in Cnv_Settings
	rSpeedSetpoint:  REAL;                // [user units], signed
END_VAR
VAR_TEMP
	Execute_Old:  BOOL;
	Stop_Old:  BOOL;
	Forward:  Bool;
	Backward:  Bool;
	SftyPinUp:  Bool;
	SftyPinDown:  BOOL;
END_VAR

R_Start_DB(CLK := Cnv_Control.Instruction.Execute AND NOT Execute_Old);
R_Stop_DB(CLK := Cnv_Control.Instruction.Stop AND NOT Stop_Old);

Execute_Old := Cnv_Control.Instruction.Execute;
Stop_Old := Cnv_Control.Instruction.Stop;

Cnv_Control.Enabled := Cnv_Control.Instruction.Enable OR Cnv_Control.Mode = 3;

ID_Decode_F(ID := Cnv_Settings.ID,
            ID_Decoded := ID_Decoded);

ID_Decode_F(ID := Cnv_Control.Instruction.Transfer_From_ID,
              ID_Decoded := ID_Decoded_From);

ID_Decode_F(ID := Cnv_Control.Instruction.Transfer_To_ID,
              ID_Decoded := ID_Decoded_To);

//MODES
Cnv_Control.Mode := Cnv_Control.Instruction.Mode_Change;
IF (Cnv_Control.Mode = 1 OR Cnv_Control.Mode = 5) AND NOT Cnv_Control.Error THEN
    State := 500;
END_IF;

R_Automatic_Mode(CLK := Cnv_Control.Mode = 3);
IF R_Automatic_Mode.Q OR (NOT Cnv_Control.Enabled AND NOT Cnv_Control.Error) THEN
    State := 0;
END_IF;

(*
Mode select is done via the HMI. Might add external mode select switches.
        
        Mode select mask:
        0: Disabled
        1: Manual
        2: Semi-Auto
        3: Auto
        4: Teach - N/A for Cnv
        5: Maintenance
        
Device ID Format: XXYYZZ    
XX = Device type   
    40  VTD
    10  Cnv_Front_of_VTD
    11  Cnv_Rear_of_VTD
    12  Cnv_On_Extractor
	13  Turn_Table
    20  Safety_Stop_Front_of_VTD
    21  Safety_Stop_Rear_of_VTD
  
YY = Floor   
ZZ = VTD Connected to    
Example: 110203 Conveyor at the rear of VTD 3 on level 2    
*)

{region "Sensor allocations"}
    //PALLET DETECT
    Forward := Cnv_Control.Inputs.Forward_Sensor;
    Backward := Cnv_Control.Inputs.Backward_Sensor;
    
    //SAFETY PINS (IT DOESN'T EXIST IN ECONVEYORS)
    SftyPinUp := Cnv_Control.Safety_Stop_Cnrl.Inputs.DP_Extended;
    SftyPinDown := Cnv_Control.Safety_Stop_Cnrl.Inputs.DP_Retracted;
{endregion}

{region "Cyclic Checks"}
    // Check Pallet
    T_CheckPallet(IN:=Forward AND Backward,
                   PT:=Time_CheckPallet);
    
    T_CheckNoPallet(IN:=Cnv_Control.Running AND NOT Forward AND NOT Backward,
                   PT:=Time_CheckNoPallet);
    
    //Conditions for Conveyor occupied
  IF T_CheckPallet.Q OR // Both sensors triggered after a timer
        (NOT Forward AND Backward AND NOT Cnv_Control.Running) OR //Forward sensor triggered and not running
        (Forward AND NOT Backward AND NOT Cnv_Control.Running) //Backward sensor triggered and not running
    THEN
        Cnv_Control.Cnv_Occupied := TRUE;//Conveyor occupied
    ELSIF T_CheckNoPallet.Q OR //Check pallet Timer
        (NOT Cnv_Control.Running AND NOT Forward AND NOT Backward) //No sensor detected and Conveyor not running
    THEN
        //No Pallet
        Cnv_Control.Cnv_Occupied := FALSE;
    END_IF;
    
    // Update the Cnv_Control opbject
    Cnv_Control.SM_State := State;
    Cnv_Control.Stopped := NOT Cnv_Control.Running;
    IF Cnv_Control.Instruction.Inbound_Ready OR Cnv_Control.Instruction.Outbound_Ready THEN
        Cnv_Control.Ready_For_Task := TRUE;
    ELSE
        Cnv_Control.Ready_For_Task := FALSE;
    END_IF;
    
    IF ID_Decoded.Device_Type = 10 THEN
        Settings.LCnv[ID_Decoded.Level].Cnv_Level := INT_TO_UINT(ID_Decoded.Level);
    END_IF;
{endregion}

{region "Auto/Semi auto mode"}
    CASE State OF
        0: //Initialization
            Cnv_Control.Instruction.Inbound_Ready := FALSE;
            Cnv_Control.Instruction.Outbound_Ready := FALSE;
            Cnv_Control.Instruction.Transfer_Complete := FALSE;
            Cnv_Control.Instruction.Transfer_in_Progress := FALSE;
            Cnv_Control.Running := FALSE;
            Cnv_Control.Motor.Forward := FALSE;
            Cnv_Control.Motor.Reverse := FALSE;
            Cnv_Control.Motor.Speed := 0;
            Timer_Transfer(IN := FALSE,
                            PT := T#0S);
            T_Ramp(IN := FALSE,
                    PT := t#0s);
            IF Cnv_Control.Enabled AND (Cnv_Control.Mode = 3 OR Cnv_Control.Mode = 2) AND NOT Cnv_Control.Error THEN
                State := 10;
            END_IF;
            
        10: //Standby - Conveyor ready to receive instruction
            IF Cnv_Control.Ready_For_Task AND (R_Start_DB.Q OR Cnv_Control.Instruction.Start_Transfer)
            THEN //WCS NORMAL TRANSFER
                Cnv_Control.Instruction.Inbound_Ready := FALSE;
                Cnv_Control.Instruction.Outbound_Ready := FALSE;
                Cnv_Control.Done := FALSE;
                Cnv_Control.Running := TRUE;
                Cnv_Control.Instruction.Transfer_in_Progress := TRUE;
                Cnv_Control.Current_Task_ID := Cnv_Control.Instruction.Task_ID;
                State := 20;
            ELSIF Cnv_Control.Instruction.Start_Transfer AND ID_Decoded.Level = 10 AND VTD_Level <> Cnv_Settings.Cnv_Level THEN
                //Extractor not at the correct level
                Set_Bit_F(BIT_Number := 2,
                            Variavel := Cnv_Control.Cnv_Errors.Error_Word_3);
            END_IF;
            
            //----------------------- Pallet Movement -----------------------
        20: //Set the direction of transfer
            IF ID_Decoded.Device_Type = 10 AND ID_Decoded_From.Device_Type = 12 AND NOT Cnv_Control.Cnv_Occupied AND
                Control.ECnv.Cnv_Occupied THEN //Extractor to CNV 1
                Cnv_Control.Motor.Speed := Cnv_Settings.Full_Speed;
                Cnv_Control.Motor.Forward := TRUE;
                Transfer_Direction := 'Forward';
                State := 30;
            ELSIF ID_Decoded.Device_Type = 10 AND ID_Decoded_To.Device_Type = 12 AND Cnv_Control.Cnv_Occupied AND
                NOT Control.ECnv.Cnv_Occupied THEN //CNV 1 To extractor
                IF Control.ECnv.SM_State = 30 THEN //Wait CVTD RUn
                    Cnv_Control.Motor.Speed := Cnv_Settings.Full_Speed;
                    Cnv_Control.Motor.Reverse := TRUE;
                    Transfer_Direction := 'Backward';
                    State := 30;
                END_IF;
            ELSE //14:3 Cnv cannot transfer to that location
                Set_Bit_F(BIT_Number := 5,
                            Variavel := Cnv_Control.Cnv_Errors.Error_Word_2);
            END_IF;
            
        30: // Running
            IF R_Stop_DB.Q THEN
                Cnv_Control.Motor.Forward := FALSE;
                Cnv_Control.Motor.Reverse := FALSE;
                Cnv_Control.Motor.Speed := 0;
                State := 0;
            ELSE
                //Slowdown ramp
                T_Ramp(IN := TRUE,
                        PT := Time_SlowDown_Ramp);
                IF T_Ramp.ET > (Time_SlowDown_Ramp * 70) / 100 AND T_Ramp.ET < (Time_SlowDown_Ramp * 80) / 100 THEN
                    Cnv_Control.Motor.Speed := Cnv_Settings.Slow_Speed * 3;
                ELSIF T_Ramp.ET > (Time_SlowDown_Ramp * 80) / 100 AND T_Ramp.ET < (Time_SlowDown_Ramp * 90) / 100 THEN
                    Cnv_Control.Motor.Speed := Cnv_Settings.Slow_Speed * 2;
                ELSIF T_Ramp.ET >= Time_SlowDown_Ramp THEN
                    Cnv_Control.Motor.Speed := Cnv_Settings.Slow_Speed;
                END_IF;
            END_IF;
            
            //Check conditions to stop the motor
            IF (ID_Decoded.Device_Type = 10 AND ID_Decoded_From.Device_Type = 12) //ECONV To CNV 1 - 10(CNV1)
            THEN
                IF Cnv_Control.Cnv_Occupied THEN //Stop the motor if the conveyor is not occupied anymore
                    State := 35;
                END_IF;
            ELSIF (ID_Decoded.Device_Type = 10 AND ID_Decoded_To.Device_Type = 12) //CNV 1 To ECNV - 10(CNV1)
            THEN
                IF NOT Cnv_Control.Cnv_Occupied THEN //Stop the motor if the conveyor is occupied
                    State := 35;
                END_IF;
            END_IF;
            
            //Monitor the transfer progress
            Timer_Transfer(IN := TRUE,
                            PT := UINT_TO_TIME(Cnv_Settings.Transfer_Time) * 1000);
            //If the watchdog bites, kill the process
            IF Timer_Transfer.Q THEN //14:1 Transfer timed out
                Set_Bit_F(BIT_Number := 3,
                           Variavel := Cnv_Control.Cnv_Errors.Error_Word_2);
            END_IF;
            
        35: //Stop motor
                T_Ramp(IN := FALSE,
                        PT := T#0S);
                Cnv_Control.Motor.Forward := FALSE;
                Cnv_Control.Motor.Reverse := FALSE;
                Cnv_Control.Motor.Speed := 0;
                Cnv_Control.Done := TRUE;
                State := 0;
            
        //----------------------- Pallet Alignment -----------------------
        400: //Error state
            Cnv_Control.Instruction.Inbound_Ready := FALSE;
            Cnv_Control.Instruction.Outbound_Ready := FALSE;
            Cnv_Control.Running := FALSE;
            Cnv_Control.Motor.Speed := 0;
            Cnv_Control.Motor.Forward := FALSE;
            Cnv_Control.Motor.Reverse := FALSE;
            Cnv_Control.Instruction.Stop := FALSE;
            Cnv_Control.Instruction.Transfer_in_Progress := FALSE;
            Watchdog(IN := FALSE,
                      PT := T#0S);
            Timer_Transfer(IN := FALSE,
                            PT := T#0S);

            T_Ramp(IN := FALSE,
                    PT := t#0s);
            IF Cnv_Control.Instruction.Reset OR SYSTEM_CONTROL.Reset_All OR HMI_Reset THEN
                Cnv_Control.Warning := 0;
                Cnv_Control.Current_Task_ID := 0;
                Cnv_Control.Error := FALSE; //Reset the conveyor
                
                Cnv_Control.Cnv_Errors.Error_Word_1 := 0;
                Cnv_Control.Cnv_Errors.Error_Word_2 := 0;
                Cnv_Control.Cnv_Errors.Error_Word_3 := 0;
                Cnv_Control.Cnv_Errors.Error_Word_4 := 0;
                State := 0;
            END_IF;
            
        500:
            IF Cnv_Control.Enabled THEN
                IF Cnv_Control.Instruction.Foward OR
                    (ID_Decoded.Device_Type = 10 AND Cnv_Control.Instruction.Start_Transfer AND NOT CNV_In_Out AND CNV1_2_Selected = 1 (*RECEIVE = 0*)) OR
                    (ID_Decoded.Device_Type = 10 AND Cnv_Control.Instruction.Start_Transfer AND CNV_In_Out AND CNV1_2_Selected = 2 (*SEND = 1*))
                THEN
                    Cnv_Control.Motor.Speed := Cnv_Settings.Manual_Speed;
                    Cnv_Control.Motor.Forward := TRUE;
                    Cnv_Control.Running := TRUE;
                ELSIF Cnv_Control.Instruction.Backward OR
                    (ID_Decoded.Device_Type = 10 AND Cnv_Control.Instruction.Start_Transfer AND NOT CNV_In_Out AND CNV1_2_Selected = 2 (*RECEIVE = 0*)) OR
                    (ID_Decoded.Device_Type = 10 AND Cnv_Control.Instruction.Start_Transfer AND CNV_In_Out AND CNV1_2_Selected = 1 (*SEND = 1*))
                THEN
                    Cnv_Control.Motor.Speed := Cnv_Settings.Manual_Speed;
                    Cnv_Control.Motor.Reverse := TRUE;
                    Cnv_Control.Running := TRUE;
                ELSE
                    Cnv_Control.Motor.Speed := 0;
                    Cnv_Control.Motor.Forward := FALSE;
                    Cnv_Control.Motor.Reverse := FALSE;
                    Cnv_Control.Running := FALSE;
                END_IF;
            END_IF;
            IF Cnv_Control.Mode <> 1 AND Cnv_Control.Mode <> 5 THEN
                State := 0;
            END_IF;
    END_CASE;
{endregion}

{region "Cyclic Error Checks"}
    IF NOT Safety_OK THEN //11:1
        Set_Bit_F(BIT_Number := 0,
                    Variavel := Cnv_Control.Cnv_Errors.Error_Word_1);
    END_IF;
    
    IF Cnv_Control.Motor.Error THEN
        Set_Bit_F(BIT_Number:= 0,
                  Variavel := Cnv_Control.Cnv_Errors.Error_Word_4);
    END_IF;
    
    IF Cnv_Control.Instruction.Stop THEN //HMI STOP
        Set_Bit_F(BIT_Number := 1,
                    Variavel := Cnv_Control.Cnv_Errors.Error_Word_1);
    END_IF;
    
    IF Cnv_Control.Safety_Stop_Cnrl.Error THEN
        Set_Bit_F(BIT_Number := 1,
                    Variavel := Cnv_Control.Cnv_Errors.Error_Word_4);
    END_IF;
    
    IF ((ID_Decoded.VTD = 1 AND ERRORS.Errors_Profinet_1.8) OR
        (ID_Decoded.VTD = 2 AND Errors.Errors_Profinet_3.7)) AND Cnv_Control.Mode <> 1
    THEN //Profinet error
        Set_Bit_F(BIT_Number := 3,
                    Variavel := Cnv_Control.Cnv_Errors.Error_Word_3);
    END_IF;
    
    
    // go to error state
    IF Cnv_Control.Cnv_Errors.Error_Word_1 <> 0 OR
        Cnv_Control.Cnv_Errors.Error_Word_2 <> 0 OR
        Cnv_Control.Cnv_Errors.Error_Word_3 <> 0 OR
        Cnv_Control.Cnv_Errors.Error_Word_4 <> 0
    THEN
        Cnv_Control.Error := TRUE;
        State := 400;
    END_IF;
{endregion}

{region "VFD - SEW MOVIKIT Velocity Drive (5 PD)"}
    // Converted from the former G120/SinaSpeed region (kept below as SIEMENS-LEGACY comments).
    // The state machine above still commands the motor exactly as before:
    //   Cnv_Control.Motor.Forward / Reverse = direction
    //   Cnv_Control.Motor.Speed             = speed in the units of Cnv_Settings.Full/Slow/Manual_Speed
    // MOVIKIT Velocity process data: SEW manual 33959862, chapter 9 (PO/PI 1..5, mode 200 implicit).
    // Raw process data: Cnv_Control.Motor.stProcessInput (from FC Inputs) and
    // Cnv_Control.Motor.aProcessOutput (to FC Outputs).
    // ASSUMPTION (verify on the first test): Forward = negative speed setpoint, as in the
    // legacy G120 code. If the conveyor runs the wrong way, correct the direction of
    // rotation in MOVISUITE, not here.

    bDriveParamsValid := Cnv_Settings.rSewSpeedPerUnit > 0.0
                         AND Cnv_Settings.uiSewAcceleration > 0
                         AND Cnv_Settings.uiSewDeceleration > 0;

    //SETPOINT (signed, user units)
    IF Cnv_Control.Motor.Forward AND NOT Cnv_Control.Motor.Reverse THEN
        rSpeedSetpoint := -1.0 * Cnv_Control.Motor.Speed * Cnv_Settings.rSewSpeedPerUnit;
    ELSIF Cnv_Control.Motor.Reverse AND NOT Cnv_Control.Motor.Forward THEN
        rSpeedSetpoint := Cnv_Control.Motor.Speed * Cnv_Settings.rSewSpeedPerUnit;
    ELSE
        rSpeedSetpoint := 0.0;
    END_IF
    MainSetpoint := REAL_TO_INT(LIMIT(-32767.0, rSpeedSetpoint, 32767.0));

    //ENABLE / START
    bDriveMoveRequest := (Cnv_Control.Motor.Forward XOR Cnv_Control.Motor.Reverse)
                         AND MainSetpoint <> 0
                         AND bDriveParamsValid;

    // Keep the enable until the motor has stopped, so a normal stop (start = 0)
    // decelerates with the PO 4 ramp. Safety_OK or a conveyor error removes the
    // enable immediately (FCB 14 emergency stop ramp).
    bDriveEnable := Safety_OK AND NOT Cnv_Control.Error
                    AND (bDriveMoveRequest OR Cnv_Control.Motor.stStatus.bMotorTurning);

    bDriveFaultReset := Cnv_Control.Instruction.Reset OR System_Control.Reset_All OR HMI_Reset;

    fbVelocityDrive(i_stProcessInput := Cnv_Control.Motor.stProcessInput,
                    i_bEnable := bDriveEnable,
                    i_bStart := bDriveMoveRequest AND bDriveEnable,
                    i_bFaultReset := bDriveFaultReset,
                    i_iSpeedSetpoint := MainSetpoint,
                    i_uiAcceleration := Cnv_Settings.uiSewAcceleration,
                    i_uiDeceleration := Cnv_Settings.uiSewDeceleration);

    Cnv_Control.Motor.aProcessOutput := fbVelocityDrive.q_aProcessOutput;
    Cnv_Control.Motor.stStatus := fbVelocityDrive.q_stStatus;

    //Status
    Cnv_Control.Motor.Status := fbVelocityDrive.q_stStatus.wStatusWord;
    Cnv_Control.Motor.Ready := fbVelocityDrive.q_bReady;
    Cnv_Control.Motor.Enabled := fbVelocityDrive.q_stStatus.bOutputStageEnabled;
    // Drive error, communication error, or a move requested without valid SEW scaling.
    Cnv_Control.Motor.Error := fbVelocityDrive.q_bError
                               OR ((Cnv_Control.Motor.Forward OR Cnv_Control.Motor.Reverse) AND NOT bDriveParamsValid);

    //Actual speed, in the units of Motor.Speed (unsigned, as before)
    IF Cnv_Settings.rSewSpeedPerUnit > 0.0 THEN
        Cnv_Control.Motor.Speed_Actual := ABS(INT_TO_REAL(fbVelocityDrive.q_stStatus.iActualSpeed))
                                          / Cnv_Settings.rSewSpeedPerUnit;
    ELSE
        Cnv_Control.Motor.Speed_Actual := 0.0;
    END_IF

    //Actual torque: PI 4 is signed [0.1 % nominal motor torque]; Actual_Torque keeps the unsigned [%] format
    Cnv_Control.Motor.Actual_Torque := DINT_TO_UINT(ABS(INT_TO_DINT(fbVelocityDrive.q_stStatus.iActualTorque_0p1pct)) / 10);

    // Actual_Current is not part of the MOVIKIT Velocity 5 PD profile. It needs the
    // "additional process values of the inverter" option in MOVISUITE; not written here.
{endregion}

// SIEMENS-LEGACY: former G120/SinaSpeed region, replaced by the region above.
// SIEMENS-LEGACY: {REGION VFD}
// SIEMENS-LEGACY:     //Status
// SIEMENS-LEGACY:     Cnv_Control.Motor.Ready := (Cnv_Control.Inputs.VFD_Status.%X0 OR Cnv_Control.Inputs.VFD_Status.%X1) AND NOT Cnv_Control.Motor.Error;
// SIEMENS-LEGACY:     Cnv_Control.Motor.Error := Cnv_Control.Inputs.VFD_Status.%X3 OR Cnv_Control.Inputs.VFD_Status.%X7 OR NOT Cnv_Control.Inputs.VFD_Status.%X13;
// SIEMENS-LEGACY:     Cnv_Control.Motor.Enabled := Cnv_Control.Inputs.VFD_Status.%X2;
// SIEMENS-LEGACY:     Cnv_Control.Motor.Actual_Current := SCALE_X(MIN := 0,
// SIEMENS-LEGACY:                                                  VALUE := NORM_X(MIN := 0,
// SIEMENS-LEGACY:                                                                  VALUE := Cnv_Control.Inputs.VFD_ActualCurrent,
// SIEMENS-LEGACY:                                                                  MAX := 16384),
// SIEMENS-LEGACY:                                                  MAX := 1.98);
// SIEMENS-LEGACY:
// SIEMENS-LEGACY:
// SIEMENS-LEGACY:     //Actual Speed
// SIEMENS-LEGACY:     IF MainSetpoint > 0 THEN
// SIEMENS-LEGACY:         Cnv_Control.Motor.Speed_Actual := SCALE_X(MIN := 0,
// SIEMENS-LEGACY:                                                    VALUE := NORM_X(MIN := 0,
// SIEMENS-LEGACY:                                                                    VALUE := Cnv_Control.Inputs.VFD_Speed_Actual,
// SIEMENS-LEGACY:                                                                    MAX := 16384),
// SIEMENS-LEGACY:                                                    MAX := 130);
// SIEMENS-LEGACY:
// SIEMENS-LEGACY:         Cnv_Control.Motor.Actual_Torque := SCALE_X(MIN := 0,
// SIEMENS-LEGACY:                                                     VALUE := NORM_X(MIN := 0,
// SIEMENS-LEGACY:                                                                     VALUE := Cnv_Control.Inputs.VFD_ActualTorque,
// SIEMENS-LEGACY:                                                                     MAX := 16384),
// SIEMENS-LEGACY:                                                     MAX := 100);
// SIEMENS-LEGACY:     ELSIF MainSetpoint < 0 THEN
// SIEMENS-LEGACY:         Cnv_Control.Motor.Speed_Actual := SCALE_X(MIN := 0,
// SIEMENS-LEGACY:                                                    VALUE := NORM_X(MIN := 0,
// SIEMENS-LEGACY:                                                                    VALUE := Cnv_Control.Inputs.VFD_Speed_Actual * -1,
// SIEMENS-LEGACY:                                                                    MAX := 16384),
// SIEMENS-LEGACY:                                                    MAX := 130);
// SIEMENS-LEGACY:
// SIEMENS-LEGACY:         Cnv_Control.Motor.Actual_Torque := SCALE_X(MIN := 0,
// SIEMENS-LEGACY:                                                     VALUE := NORM_X(MIN := 0,
// SIEMENS-LEGACY:                                                                     VALUE := Cnv_Control.Inputs.VFD_ActualTorque * -1,
// SIEMENS-LEGACY:                                                                     MAX := 16384),
// SIEMENS-LEGACY:                                                     MAX := 100);
// SIEMENS-LEGACY:     ELSE
// SIEMENS-LEGACY:         Cnv_Control.Motor.Speed_Actual := 0;
// SIEMENS-LEGACY:         Cnv_Control.Motor.Actual_Torque := 0;
// SIEMENS-LEGACY:     END_IF;
// SIEMENS-LEGACY:
// SIEMENS-LEGACY:     //MAIN SETPOINT
// SIEMENS-LEGACY:     IF Cnv_Control.Motor.Forward THEN
// SIEMENS-LEGACY:         MainSetpoint := (SCALE_X(MIN := 0,
// SIEMENS-LEGACY:                                   VALUE := NORM_X(MIN := 0,
// SIEMENS-LEGACY:                                                   VALUE := Cnv_Control.Motor.Speed (** 1.681*),
// SIEMENS-LEGACY:                                                   MAX := 130),
// SIEMENS-LEGACY:                                   MAX := 1865.0) * -1);
// SIEMENS-LEGACY:     ELSIF Cnv_Control.Motor.Reverse THEN
// SIEMENS-LEGACY:         MainSetpoint := SCALE_X(MIN := 0,
// SIEMENS-LEGACY:                                  VALUE := NORM_X(MIN := 0,
// SIEMENS-LEGACY:                                                  VALUE := Cnv_Control.Motor.Speed (** 1.681*),
// SIEMENS-LEGACY:                                                  MAX := 130),
// SIEMENS-LEGACY:                                  MAX := 1865.0);
// SIEMENS-LEGACY:     ELSE
// SIEMENS-LEGACY:         MainSetpoint := 0;
// SIEMENS-LEGACY:     END_IF;
// SIEMENS-LEGACY:
// SIEMENS-LEGACY:     SinaSpeed(EnableAxis := Cnv_Control.Motor.Forward OR Cnv_Control.Motor.Reverse,
// SIEMENS-LEGACY:                AckError := Cnv_Control.Instruction.Reset OR "Reset_All" OR HMI_Reset,
// SIEMENS-LEGACY:                SpeedSp := MainSetpoint,
// SIEMENS-LEGACY:                RefSpeed := 1865.0,
// SIEMENS-LEGACY:                HWIDSTW := Cnv_Settings.G120_Hardware_ID,
// SIEMENS-LEGACY:                HWIDZSW := Cnv_Settings.G120_Hardware_ID);
// SIEMENS-LEGACY: {END_REGION}

// TODO: HMI reset. The Siemens screen DBs below have no TwinCAT equivalent yet;
//       HMI_Reset stays FALSE until the conveyor HMI interface (GVL_HMI_*) exists.
// SIEMENS-LEGACY: HMI_Reset := "Screen_DB_1".Reset_All[1] OR "Screen_DB_1".Reset_All[2] OR "CNV_HMI"."Reset(1)"[1] OR "CNV_HMI"."Reset(1)"[2];
;

END_FUNCTION_BLOCK

// ---- POUs/SEW/FB_SEW_VelocityDrive.TcPOU
// Communication and status layer for a SEW drive running MOVIKIT Velocity
// with the "5 PD" basic process data profile (SBusPLUS, not CiA402).
// Source: SEW manual 33959862 "MOVIKIT Positioning, Velocity", chapter 4.2
// and chapter 9 "Process data assignment". Only words and bits marked V/P
// (available with MOVIKIT Velocity) are used.
//
// MOVIKIT Velocity always runs operating mode Speed (200): there is no PO 6.
// PO 1 control word, PO 2 setpoint speed, PO 3 acceleration, PO 4 deceleration,
// PO 5 digital outputs. PI 1 status word, PI 2 actual speed, PI 3 fault/subfault,
// PI 4 torque, PI 5 digital inputs.
//
// This block does NOT decide any motion. The owner of the axis (e.g.
// Buffer_Conveyor_FB) sets the commands; this block only packs them into
// PO 1..5, decodes PI 1..5 and supervises the communication
// (EtherCAT state + MOVIKIT handshake).
//
// Safety-related behavior:
//  - Enable and start are forced to 0 while communication is not OK.
//  - PO 1.3 "Release brake (without enable)" is never set.
//  - PO 1.13 "Output stage inhibit" is never set; removing enable stops the
//    drive with the emergency stop ramp (FCB 14).
FUNCTION_BLOCK FB_SEW_VelocityDrive
VAR_INPUT
    i_stProcessInput : ST_SEW_ProcessInput5;  // Raw PI 1..5 + EtherCAT diagnostics (from FC Inputs)

    i_bEnable : BOOL;                         // PO 1.0 + PO 1.1 enable (FALSE = stop with FCB 14)
    i_bStart : BOOL;                          // PO 1.7 start/stop with fieldbus ramp
    i_bFaultReset : BOOL;                     // PO 1.8, drive resets on the rising edge

    i_iSpeedSetpoint : INT;                   // PO 2, signed, user units
    i_uiAcceleration : UINT;                  // PO 3, user units
    i_uiDeceleration : UINT;                  // PO 4, user units

    i_tHandshakeTimeout : TIME := T#1S;       // Max time for PI 1.15 to follow PO 1.15
END_VAR
VAR_OUTPUT
    q_aProcessOutput : ARRAY[1..5] OF UINT;   // Raw PO 1..5 (to FC Outputs)
    q_stStatus : ST_SEW_VelocityStatus;       // Decoded PI 1..5

    q_bReady : BOOL;                          // Communication OK, ready, STO inactive, no error
    q_bError : BOOL;                          // Drive error or communication error
    q_udiErrorId : UDINT;                     // See ERROR_ID_* below, or PI 3 (fault * 256 + subfault)
END_VAR
VAR
    bHandshakeIn : BOOL;                      // Value sent in PO 1.15
    bHandshakeWaiting : BOOL;
    tonHandshake : TON;
    wControlWord : WORD;
END_VAR
VAR CONSTANT
    ERROR_ID_ETHERCAT : UDINT := 16#FFFF0001; // Drive not in OP or working counter invalid
    ERROR_ID_HANDSHAKE : UDINT := 16#FFFF0002; // MOVIKIT handshake timeout
END_VAR

{region "Communication supervision"}
// EtherCAT: state OP (lower nibble = 8) and valid working counter.
q_stStatus.bEtherCatOk := (NOT i_stProcessInput.bWcStateError)
                          AND ((i_stProcessInput.uiEcState AND 16#000F) = 8);

// MOVIKIT handshake (manual chapter 9.3): the drive copies PO 1.15 to PI 1.15.
// When both are equal, invert PO 1.15; otherwise the timeout runs.
q_stStatus.bHandshakeOut := i_stProcessInput.aWord[1].15;

IF q_stStatus.bEtherCatOk THEN
    IF bHandshakeIn = q_stStatus.bHandshakeOut THEN
        bHandshakeIn := NOT bHandshakeIn;
        bHandshakeWaiting := FALSE;
    ELSE
        bHandshakeWaiting := TRUE;
    END_IF
ELSE
    // No valid data: the EtherCAT error is reported instead of the handshake.
    bHandshakeWaiting := FALSE;
END_IF

tonHandshake(IN := bHandshakeWaiting, PT := i_tHandshakeTimeout);
q_stStatus.bHandshakeError := tonHandshake.Q;

q_stStatus.bCommunicationOk := q_stStatus.bEtherCatOk AND NOT q_stStatus.bHandshakeError;
{endregion}

{region "Decode process inputs (PI 1..5)"}
q_stStatus.wStatusWord := UINT_TO_WORD(i_stProcessInput.aWord[1]);
q_stStatus.bReady := q_stStatus.wStatusWord.0;
q_stStatus.bStoInactive := q_stStatus.wStatusWord.1;
q_stStatus.bOutputStageEnabled := q_stStatus.wStatusWord.2;
q_stStatus.bBrakeReleased := q_stStatus.wStatusWord.3;
q_stStatus.bMotorTurning := q_stStatus.wStatusWord.4;
q_stStatus.bError := q_stStatus.wStatusWord.8;
q_stStatus.bWarning := q_stStatus.wStatusWord.9;
q_stStatus.bDriveTrain2Active := q_stStatus.wStatusWord.10;
q_stStatus.bSpeedReached := q_stStatus.wStatusWord.11;
q_stStatus.bStandbyActive := q_stStatus.wStatusWord.14;
// Bits 5, 6, 7 and 12 exist only with MOVIKIT Positioning and are not decoded.

// Same-size integer conversions keep the bit pattern (signed values).
q_stStatus.iActualSpeed := UINT_TO_INT(i_stProcessInput.aWord[2]);
q_stStatus.byFaultCode := WORD_TO_BYTE(SHR(UINT_TO_WORD(i_stProcessInput.aWord[3]), 8));
q_stStatus.bySubfaultCode := WORD_TO_BYTE(UINT_TO_WORD(i_stProcessInput.aWord[3]) AND 16#00FF);
q_stStatus.iActualTorque_0p1pct := UINT_TO_INT(i_stProcessInput.aWord[4]);
q_stStatus.wDigitalInputs := UINT_TO_WORD(i_stProcessInput.aWord[5]);
{endregion}

{region "Diagnostics"}
q_bError := q_stStatus.bError OR NOT q_stStatus.bCommunicationOk;
q_bReady := q_stStatus.bCommunicationOk AND q_stStatus.bReady
            AND q_stStatus.bStoInactive AND NOT q_stStatus.bError;

IF NOT q_stStatus.bEtherCatOk THEN
    q_udiErrorId := ERROR_ID_ETHERCAT;
ELSIF q_stStatus.bHandshakeError THEN
    q_udiErrorId := ERROR_ID_HANDSHAKE;
ELSIF q_stStatus.bError THEN
    q_udiErrorId := UINT_TO_UDINT(i_stProcessInput.aWord[3]);
ELSE
    q_udiErrorId := 0;
END_IF
{endregion}

{region "Build process outputs (PO 1..5)"}
wControlWord := 0;

IF q_stStatus.bCommunicationOk AND i_bEnable THEN
    wControlWord.0 := TRUE;     // Enable/emergency stop
    wControlWord.1 := TRUE;     // Enable/application stop
    wControlWord.7 := i_bStart; // Start/stop with fieldbus ramp
END_IF

wControlWord.8 := i_bFaultReset;  // Allowed without enable
wControlWord.15 := bHandshakeIn;  // MOVIKIT handshake, no effect on motion
// Never set: bit 3 (release brake without enable), bit 10 (drive train 2),
// bit 13 (output stage inhibit), bit 14 (standby).
// Bits 4, 5, 6 and 12 exist only with MOVIKIT Positioning.

q_aProcessOutput[1] := WORD_TO_UINT(wControlWord);

IF q_stStatus.bCommunicationOk AND i_bEnable THEN
    q_aProcessOutput[2] := INT_TO_UINT(i_iSpeedSetpoint);
ELSE
    q_aProcessOutput[2] := 0;
END_IF

q_aProcessOutput[3] := i_uiAcceleration;
q_aProcessOutput[4] := i_uiDeceleration;
q_aProcessOutput[5] := 0;  // Drive digital outputs not used
{endregion}

END_FUNCTION_BLOCK

// ---- POUs/System/Functions/ID_Decode_F.TcPOU
FUNCTION ID_Decode_F : BOOL
VAR_INPUT
    ID : DINT;
END_VAR
VAR_IN_OUT
    ID_Decoded : ID_Decoded_DUT;
END_VAR

// Source: Reference_Project/ID_Decode_F.scl. Decimal layout: XXYYZZ.
// Zero is accepted as the unassigned ID. Reject negative or oversized IDs.
ID_Decode_F := FALSE;
ID_Decoded.Device_Type := 0;
ID_Decoded.Level := 0;
ID_Decoded.VTD := 0;
IF (ID < DINT#0) OR (ID > DINT#999999) THEN
    RETURN;
END_IF;
ID_Decoded.Device_Type := DINT_TO_INT(ID / DINT#10000);
ID_Decoded.Level := DINT_TO_INT((ID MOD DINT#10000) / DINT#100);
ID_Decoded.VTD := DINT_TO_INT(ID MOD DINT#100);
ID_Decode_F := TRUE;

END_FUNCTION

// ---- POUs/System/Functions/Set_Bit_F.TcPOU
FUNCTION Set_Bit_F : BOOL
VAR_INPUT
    BIT_Number : UINT;
    Bit_Value : BOOL := TRUE; // Default preserves existing set-only callers.
END_VAR
VAR_IN_OUT
    Variavel : WORD; // Existing interface name retained for compatibility.
END_VAR

// Source: Reference_Project/Set_Bit_F.scl.
// FALSE leaves the word unchanged, matching the Siemens set-only behavior.
Set_Bit_F := FALSE;
IF BIT_Number > UINT#15 THEN
    RETURN;
END_IF;
IF Bit_Value THEN
    Variavel := Variavel OR SHL(WORD#1, BIT_Number);
END_IF;
Set_Bit_F := TRUE;

END_FUNCTION

// ---- POUs/Conveyors/FB_Conveyor_MotorInterlock.TcPOU
// Grants one motor at a time inside a group of motors that must not run together
// (break-before-make). Examples: lift and transfer of a popup (inside PopUp_Conveyor_FB);
// turntable rotation and turntable roller conveyor (Control.Turn_Table.Interlock /
// Control.TBCnv.Interlock, one instance called before both device FBs).
//
// This block does NOT command any motor. The owner FB requests a motor, drives it only
// while q_abAllowed[n] is TRUE, removes Forward/Reverse as soon as the permission drops,
// and reports i_abStopped[n] (motor not turning and output stage off, from the SEW status).
// A motor whose drive communication is not OK must be reported as NOT stopped (unknown),
// so the group stays blocked until the status is valid again.
//
// Behavior:
//  - A motor is granted only when every motor of the group has been stopped for at least
//    i_tChangeover (brake closed, mechanics at rest), at start-up and at every change.
//  - The granted motor keeps the permission while its request stays TRUE.
//  - Several requests at the same time: the lowest index wins.
//  - i_iMotorCount outside 1..4 or i_tChangeover = T#0S: not configured, nothing is granted.
//  - Drive status is the owner's value of the previous cycle: one PLC cycle delay.
//
// Diagnostics:
//  - q_bConflict: more than one motor of the group is not stopped. Should never happen;
//    the owner must stop its motors and report an error.
//
// Functional interlock in the standard PLC. It is NOT a safety function.
FUNCTION_BLOCK FB_Conveyor_MotorInterlock
VAR_INPUT
    i_abRequest : ARRAY[1..4] OF BOOL;      // Owner -> block: motor n wants to run
    i_abStopped : ARRAY[1..4] OF BOOL;      // Owner -> block: motor n not turning and output stage off

    i_iMotorCount : INT;                    // Motors used in this group, 1..4 (0 = not configured)
    i_tChangeover : TIME;                   // Min. time all motors are stopped before a grant (T#0S = not configured)
END_VAR
VAR_OUTPUT
    q_abAllowed : ARRAY[1..4] OF BOOL;      // Block -> owner: motor n may run

    q_iActive : INT;                        // Granted motor 1..4, 0 = none
    q_bChangeover : BOOL;                   // A motor is requested and waits for the group to be stopped
    q_bAllStopped : BOOL;                   // Every motor of the group is stopped
    q_bConflict : BOOL;                     // More than one motor of the group is not stopped
    q_bSettingsValid : BOOL;                // i_iMotorCount in 1..4 and i_tChangeover > T#0S
END_VAR
VAR
    iMotor : INT;                           // Loop index over the motors of the group
    iNotStopped : INT;                      // Number of motors not stopped
    bAnyRequest : BOOL;                     // At least one motor is requested

    tonAllStopped : TON;                    // All motors stopped for i_tChangeover
END_VAR
VAR CONSTANT
    MAX_MOTORS : INT := 4;                  // Size of the motor arrays
END_VAR

{region "Supervision"}
q_bSettingsValid := (i_iMotorCount >= 1)
                    AND (i_iMotorCount <= MAX_MOTORS)
                    AND (i_tChangeover > T#0S);

iNotStopped := 0;
bAnyRequest := FALSE;
IF q_bSettingsValid THEN
    FOR iMotor := 1 TO i_iMotorCount DO
        IF NOT i_abStopped[iMotor] THEN
            iNotStopped := iNotStopped + 1;
        END_IF
        IF i_abRequest[iMotor] THEN
            bAnyRequest := TRUE;
        END_IF
    END_FOR
END_IF

q_bAllStopped := q_bSettingsValid AND (iNotStopped = 0);
q_bConflict := (iNotStopped > 1);

// Restarts whenever a motor of the group turns.
tonAllStopped(IN := q_bAllStopped, PT := i_tChangeover);
{endregion}

{region "Release"}
// The granted motor keeps its permission only while it is requested and the group is healthy.
IF q_iActive <> 0 THEN
    IF (q_iActive < 1)
       OR (q_iActive > i_iMotorCount)
       OR NOT q_bSettingsValid
       OR q_bConflict
    THEN
        q_iActive := 0;
    ELSIF NOT i_abRequest[q_iActive] THEN
        q_iActive := 0;
    END_IF
END_IF
{endregion}

{region "Grant"}
// A new motor is granted only after every motor has been stopped for i_tChangeover.
// The loop runs downwards so that the lowest requested index wins.
IF (q_iActive = 0) AND tonAllStopped.Q THEN
    FOR iMotor := i_iMotorCount TO 1 BY -1 DO
        IF i_abRequest[iMotor] THEN
            q_iActive := iMotor;
        END_IF
    END_FOR
END_IF
{endregion}

{region "Outputs"}
FOR iMotor := 1 TO MAX_MOTORS DO
    q_abAllowed[iMotor] := (iMotor = q_iActive);
END_FOR

q_bChangeover := bAnyRequest AND (q_iActive = 0);
{endregion}

END_FUNCTION_BLOCK

// ---- POUs/DWORD_REAL.TcPOU
FUNCTION DWORD_REAL : REAL
VAR_INPUT
	b0 : BYTE;
    b1 : BYTE;
    b2 : BYTE;
    b3 : BYTE;
END_VAR
VAR
	uValue : U_DWORD_REAL1;
END_VAR

// uValue.dw :=
//     DWORD(b0)
//     OR SHL(DWORD(b1), 8)
//     OR SHL(DWORD(b2), 16)
//     OR SHL(DWORD(b3), 24);
// 
// DWORD_REAL := uValue.dw;

END_FUNCTION

// ---- POUs/Profile_Station_FC.TcPOU
FUNCTION Profile_Station_FC : BOOL
VAR_INPUT
	MaxLength : REAL;
	ConveyorSpeed_mm_s: REAL;
END_VAR
VAR
END_VAR

// "R_TRIG_DB_26"(CLK:="Control_DB"."Profiling Station".Start);
// 
//  "R_TRIG_DB_27"(CLK:=NOT "Profile Station - Cross 1" AND NOT "Profile Station - Cross 2",Q => "SensorUp");
// 
//  "IEC_Timer_0_DB_3".TON(IN:="Profile Station - Cross 1" AND "Profile Station - Cross 2",
//                         PT:=T#2s,Q=>"SensorDown");
//  
// 
// CASE "State_PS" OF
//         
//         //-------------------------------------------------
//         // 0 - IDLE
//         //-------------------------------------------------
//     0:
//         "Control_DB"."Profiling Station".Error_ID := 0;
//         "Control_DB"."Profiling Station".Ready := TRUE;
//         "Control_DB"."Profiling Station".Running := FALSE;
//         IF "R_TRIG_DB_26".Q THEN
//             "Control_DB"."Profiling Station".Ready := FALSE;
//             "Control_DB"."Profiling Station".Done := FALSE;
//             "Control_DB"."Profiling Station".Valid := FALSE;
//             "Control_DB"."Profiling Station".OverWidth := FALSE;
//             "Control_DB"."Profiling Station".OverHeight := FALSE;
//             "Control_DB"."Profiling Station".OverLength := FALSE;
//             "Control_DB"."Profiling Station".Error_ID := 0;
//             "Control_DB"."Profiling Station".Running := TRUE;
//             "State_PS" := 10;
//         END_IF;
//         
//     10:
//         IF "SensorUp" THEN
//             "State_PS" := 20;
//         END_IF;
//         
//     20:
//         "LengthTimer".TON(IN := TRUE,
//                           PT := T#60S);
//         
//         IF NOT "Profile Station - Left" OR NOT "Profile Station - Right" THEN
//             "Control_DB"."Profiling Station".OverWidth := TRUE;
//         END_IF;
//         
//         IF NOT "Profile Station - High" THEN
//             "Control_DB"."Profiling Station".OverHeight := TRUE;
//         END_IF;
//         
//         IF "SensorDown" THEN
//             "MeasuredTime_s" := DINT_TO_REAL(TIME_TO_DINT("LengthTimer".ET)) / 1000.0;
//             "CalculatedLength" := "MeasuredTime_s" * #ConveyorSpeed_mm_s;
//             
//             // IF "CalculatedLength" > #MaxLength THEN
//             //     "Control_DB"."Profiling Station".OverLength := TRUE;
//             // END_IF;
//             
//             // Resultado final
//             IF "Control_DB"."Profiling Station".OverWidth OR "Control_DB"."Profiling Station".OverHeight OR "Control_DB"."Profiling Station".OverLength THEN
//                 "Control_DB"."Profiling Station".Valid := FALSE;
//                 "Control_DB"."Profiling Station".Error_ID.%X0 := 1;
//             ELSE
//                 "Control_DB"."Profiling Station".Valid := TRUE;
//                 "Control_DB"."Profiling Station".Error_ID := 0;
//             END_IF;
//             
//             "LengthTimer".TON(IN := FALSE,
//                               PT := T#0S);
//             "State_PS" := 100;
//         END_IF;
//         
//     100:
//         "Control_DB"."Profiling Station".Running := FALSE;
//             "Control_DB"."Profiling Station".Done := TRUE;
//             "State_PS" := 0;
//             
//        
//     END_CASE;
//     
//     "IEC_Timer_0_DB_12".TON(IN:="Control_DB"."Profiling Station".Running,
//                             PT:=t#30s);
//     
//     IF "IEC_Timer_0_DB_12".Q THEN
//         "Control_DB"."Profiling Station".Valid := FALSE;
//         "Control_DB"."Profiling Station".Error_ID := 1;
//         "State_PS" := 100;
//     END_IF;
//

END_FUNCTION

// ---- POUs/Stack_Lights_FB.TcPOU
FUNCTION_BLOCK Stack_Lights_FB
VAR_INPUT
    System_Auto : BOOL;
    Fault : BOOL;
    i_bFlash_05Hz : BOOL := TRUE; // Supply a 0.5 Hz clock; otherwise fault is steady red.
END_VAR
VAR_OUTPUT
    Red : BOOL;
    Green : BOOL;
    Orange : BOOL; // Existing TwinCAT output name retained.
    Yellow : BOOL; // Source-compatible alias for Orange.
END_VAR

// Source: Reference_Project/Stack_Lights_FB.scl.
// Priority: fault, automatic, manual. Clock is explicit instead of a Siemens tag.
Red := Fault AND i_bFlash_05Hz;
Green := NOT Fault AND System_Auto;
Orange := NOT Fault AND NOT System_Auto;
Yellow := Orange;

END_FUNCTION_BLOCK

// ---- POUs/System/Barcode_Station_FB.TcPOU
FUNCTION_BLOCK Barcode_Station_FB
VAR_INPUT
    Sick_Result : STRING(254); // Complete received payload, not a physical input address.
    Reset : BOOL; // Abort the current read; does not reset the lifetime counter.
END_VAR
VAR_OUTPUT
    Counter : UINT;
END_VAR
VAR_IN_OUT
    Station_Control : Barcode_Station_DUT;
    Auto_Start_Lector : BOOL; // Request only; caller owns transport to the scanner.
    Auto_Stop_Lector : BOOL; // One-cycle stop request, not a scanner acknowledgement.
END_VAR
VAR
    State : E_BarcodeState := E_BarcodeState.Idle;
    startEdge : R_TRIG;
    readTimer : TON;
    gateNumber : STRING(254);
    readingGateCount : STRING(254);
    code : STRING(254);
END_VAR

// Adapted from Reference_Project/Barcode_Station_FB.scl.
// No device or network mapping is performed by this block.
startEdge(CLK := Station_Control.Start);
readTimer(IN := (State = E_BarcodeState.Reading) AND NOT Reset, PT := T#15S);
Auto_Start_Lector := FALSE;
Auto_Stop_Lector := FALSE;

IF Reset THEN
    Auto_Stop_Lector := State <> E_BarcodeState.Idle;
    State := E_BarcodeState.Idle;
    Station_Control.Start := FALSE;
    Station_Control.Ready := TRUE;
    Station_Control.Running := FALSE;
    Station_Control.Done := FALSE;
    Station_Control.Valid := FALSE;
    Station_Control.Barcode := '';
    RETURN;
END_IF;

CASE State OF
    E_BarcodeState.Idle:
        Station_Control.Ready := TRUE;
        Station_Control.Running := FALSE;
        IF startEdge.Q THEN
            Station_Control.Start := FALSE;
            Station_Control.Ready := FALSE;
            Station_Control.Running := TRUE;
            Station_Control.Done := FALSE;
            Station_Control.Valid := FALSE;
            Station_Control.Barcode := '';
            // Ignore an already-present result from the preceding scan transaction.
            Station_Control.Reading_Gate_number_OLD := FindStringField(
                FieldName := 'Number', JsonStr := Sick_Result);
            State := E_BarcodeState.Reading;
        END_IF;

    E_BarcodeState.Reading:
        Station_Control.Start := FALSE;
        Station_Control.Ready := FALSE;
        Station_Control.Running := TRUE;
        Auto_Start_Lector := TRUE;
        gateNumber := FindStringField(FieldName := 'Number', JsonStr := Sick_Result);
        readingGateCount := FindStringField(FieldName := 'NRG', JsonStr := Sick_Result);
        code := FindStringField(FieldName := 'Code', JsonStr := Sick_Result);
        Station_Control.Reading_Gate_number := gateNumber;
        Station_Control.Number_OF_Reading_Gates := readingGateCount;
        Station_Control.Number_OF_Reading_Gates_OLD := readingGateCount;

        IF ((gateNumber <> '') AND
            (gateNumber <> Station_Control.Reading_Gate_number_OLD)) OR readTimer.Q THEN
            Auto_Start_Lector := FALSE;
            Station_Control.Valid := (gateNumber <> '') AND
                (gateNumber <> Station_Control.Reading_Gate_number_OLD) AND (code <> '');
            IF Station_Control.Valid THEN
                Station_Control.Barcode := code;
                Station_Control.Barcode_Old := code;
            ELSE
                Station_Control.Barcode := '';
            END_IF;
            IF gateNumber <> '' THEN
                Station_Control.Reading_Gate_number_OLD := gateNumber;
            END_IF;
            State := E_BarcodeState.Complete;
        END_IF;

    E_BarcodeState.Complete:
        Auto_Stop_Lector := TRUE;
        IF Counter = UINT#65535 THEN
            Counter := 0;
        ELSE
            Counter := Counter + 1;
        END_IF;
        Station_Control.Running := FALSE;
        Station_Control.Done := TRUE;
        Station_Control.Ready := FALSE;
        State := E_BarcodeState.Idle;

ELSE
    // Recover deterministically from an invalid state without accepting a result.
    Auto_Stop_Lector := TRUE;
    Station_Control.Start := FALSE;
    Station_Control.Running := FALSE;
    Station_Control.Ready := FALSE;
    Station_Control.Done := FALSE;
    Station_Control.Valid := FALSE;
    Station_Control.Barcode := '';
    State := E_BarcodeState.Idle;
END_CASE;

END_FUNCTION_BLOCK

// ---- POUs/System/Functions/FindStringField.TcPOU
FUNCTION FindStringField : STRING(254)
VAR_INPUT
    FieldName : STRING(254);
    JsonStr : STRING(254);
END_VAR
VAR
    pattern : STRING(254);
    character : STRING(1);
    foundPos : INT;
    cursor : INT;
    valueStart : INT;
    length : INT;
    scan : INT;
END_VAR

// Adapted from Reference_Project/Barcode_Station_FB.scl.
// Extract a plain quoted field from the flat SICK payload format.
// Whitespace around ':' is accepted. Escaped values are rejected.
// This is not a general-purpose JSON validator or MQTT parser.
FindStringField := '';
IF (LEN(FieldName) = 0) OR (LEN(FieldName) > 250) THEN
    RETURN;
END_IF;
pattern := CONCAT('"', FieldName);
pattern := CONCAT(pattern, '"');
foundPos := FIND(JsonStr, pattern);
IF foundPos = 0 THEN
    RETURN;
END_IF;
length := LEN(JsonStr);
cursor := foundPos + LEN(pattern);
// Skip JSON whitespace before the colon, with a bounded scan.
FOR scan := cursor TO length DO
    character := MID(JsonStr, 1, scan);
    IF (character <> ' ') AND (character <> '$T') AND
       (character <> '$R') AND (character <> '$N') THEN
        EXIT;
    END_IF;
END_FOR;
IF scan > length THEN
    RETURN;
END_IF;
IF MID(JsonStr, 1, scan) <> ':' THEN
    RETURN;
END_IF;
cursor := scan + 1;
FOR scan := cursor TO length DO
    character := MID(JsonStr, 1, scan);
    IF (character <> ' ') AND (character <> '$T') AND
       (character <> '$R') AND (character <> '$N') THEN
        EXIT;
    END_IF;
END_FOR;
IF scan > length THEN
    RETURN;
END_IF;
IF MID(JsonStr, 1, scan) <> '"' THEN
    RETURN;
END_IF;
valueStart := scan + 1;
FOR scan := valueStart TO length DO
    character := MID(JsonStr, 1, scan);
    IF (character = '$5C') OR (character = '$R') OR
       (character = '$N') OR (character = '$T') THEN
        RETURN;
    END_IF;
    IF character = '"' THEN
        IF scan > valueStart THEN
            FindStringField := MID(JsonStr, scan - valueStart, valueStart);
        END_IF;
        RETURN;
    END_IF;
END_FOR;

END_FUNCTION

// ---- POUs/System/Conveyors_Transfer.TcPOU
FUNCTION Conveyors_Transfer : BOOL
VAR_INPUT
END_VAR
VAR
	i_Lev:  UINT;
	Concat1:  String;
	Concat2:  String;
	ID:  DInt;
	StrLev:  String;
	StrSys:  String;
	Level:  UINT;
END_VAR

StrSys := '1'; // SpaceX Inbound has one VTD system: the ID suffix stays 1

{region "ID OF THE VTD CONVEYOR"}
    FOR i_Lev := Settings.VTD.Lowest_Level TO Settings.VTD.Highest_Level DO
        IF Control.VTD.Current_Level = i_Lev THEN
            StrLev := UINT_TO_STRING(i_Lev);
            
            // Remove "+"
            IF StrLev[1] = '+' THEN
                StrLev := RIGHT(StrLev, L := LEN(StrLev) - 1);
            END_IF;
            
            //Build ID
            Concat1 := CONCAT('120', StrLev);
            Concat2 := CONCAT(Concat1, '0');
            ID := STRING_TO_DINT(CONCAT(Concat2, StrSys));
            
            Settings.ECnv.ID := ID;
            Settings.ECnv.Cnv_Level := i_Lev;
        END_IF;
    END_FOR;
{endregion}
    
{region "READY TO RECEIVE"}
    //EXTRACTOR CONVEYOR
    FOR i_Lev := 2 TO Settings.VTD.Highest_Level DO
        IF Control.VTD.Current_Level = i_Lev THEN
            StrLev := UINT_TO_STRING(i_Lev);
            
            // Remove "+"
            IF StrLev[1] = '+' THEN
                StrLev := RIGHT(StrLev, L := LEN(StrLev) - 1);
            END_IF;
            
            //Build ID
            Concat1 := CONCAT('120', StrLev);
            Concat2 := CONCAT(Concat1, '0');
            ID := STRING_TO_DINT(CONCAT(Concat2, StrSys));
        END_IF;
        
        IF Settings.ECnv.ID = ID AND NOT Control.ECnv.Error AND NOT Control.ECnv.Running
            AND NOT Control.ECnv.Cnv_Occupied AND NOT Control.ECnv.Instruction.Outbound_Ready AND
            NOT Control.LCnv[i_Lev].Running AND
            (Control.ECnv.Mode = 2 OR Control.ECnv.Mode = 3) THEN
            Control.ECnv.Instruction.Inbound_Ready := TRUE;
        END_IF;
    END_FOR;
    
    //BUFFER CONVEYORS
    FOR i_Lev := 2 TO Settings.VTD.Highest_Level DO
        //CNV 1
        IF NOT Control.LCnv[i_Lev].Error AND
            NOT Control.LCnv[i_Lev].Running AND
            NOT Control.LCnv[i_Lev].Cnv_Occupied AND
            NOT Control.LCnv[i_Lev].Instruction.Outbound_Ready AND
            (Control.LCnv[i_Lev].Mode = 2 OR Control.LCnv[i_Lev].Mode = 3) AND
            NOT Control.ECnv.Running
        THEN
            Control.LCnv[i_Lev].Instruction.Inbound_Ready := TRUE;
        END_IF;
    END_FOR;
{endregion}

{region "READY TO SEND"}
    //EXTRACTOR CONVEYOR
    Level := Settings.ECnv.Cnv_Level;
    
    IF Settings.ECnv.Cnv_Level >= 2 AND
        Settings.ECnv.Cnv_Level <= Settings.VTD.Highest_Level AND //Leveled
        Control.ECnv.Cnv_Occupied AND //Econveyor occupied
        NOT Control.ECnv.Error AND //not error
        NOT Control.ECnv.Running AND //not RUNNING
        Control.LCnv[Level].Instruction.Inbound_Ready AND 
        (Control.LCnv[Level].Mode = 2 OR
        Control.LCnv[Level].Mode = 3)  AND //cnv1 semi or auto mode
        (Control.ECnv.Mode = 2 OR Control.ECnv.Mode = 3) THEN //Econveyor semi or auto mode 
        Control.ECnv.Instruction.Outbound_Ready := TRUE;
    END_IF;
    
    
    //BUFFER CONVEYORS
    FOR i_Lev := 2 TO Settings.VTD.Highest_Level DO
        //CNV 1
        IF Control.ECnv.Instruction.Inbound_Ready AND Control.VTD.Current_Level = i_Lev AND //Extractor inbound ready
            Control.LCnv[i_Lev].Cnv_Occupied AND //Not occupied
            NOT Control.LCnv[i_Lev].Error AND NOT Control.LCnv[i_Lev].Running AND //NOT error and NOT running
            (Control.LCnv[i_Lev].Mode = 2 OR Control.LCnv[i_Lev].Mode = 3)//Semi auto or auto
        THEN 
            Control.LCnv[i_Lev].Instruction.Outbound_Ready := TRUE;
        END_IF;
    END_FOR;
{endregion}

END_FUNCTION

// ---- POUs/System/Functions/ByteArrayToString.TcPOU
FUNCTION ByteArrayToString : STRING(254)
VAR_INPUT
    Lenght : INT; // Reference spelling retained for named callers.
    ByteArray : ARRAY[0..1024] OF BYTE;
END_VAR
VAR_OUTPUT
    ByteArrayToString_1 : STRING(254);
    ByteArrayToString_2 : STRING(254);
    ByteArrayToString_3 : STRING(254);
    ByteArrayToString_4 : STRING(254);
    ByteArrayToString_5 : STRING(254);
    Truncated : BOOL;
END_VAR
VAR
    windows : ARRAY[0..5] OF STRING(254);
    window : INT;
    cursor : INT;
    first : INT;
    last : INT;
    count : INT;
    size : INT;
    skipLF : BOOL;
    value : BYTE;
END_VAR

// Six overlapping ASCII windows beginning at bytes 0,100,...,500.
// Bound input length and output capacity; no pointer copying or unbounded loops.
size := LIMIT(0, Lenght, 1025);
Truncated := (Lenght < 0) OR (Lenght > 1025) OR (size > 764);
FOR window := 0 TO 5 DO
    windows[window] := '';
    count := 0;
    skipLF := FALSE;
    first := window * 100;
    last := MIN(size - 1, first + 254);
    IF window = 5 THEN last := MIN(size - 1, 763); END_IF;
    FOR cursor := first TO last DO
        value := ByteArray[cursor];
        IF skipLF THEN
            skipLF := FALSE;
        ELSIF value <> 0 THEN
            // Match the source's removal of CRLF pairs, without removing lone CR/LF.
            IF (value = 13) AND (cursor < last) THEN
                IF ByteArray[cursor + 1] = 10 THEN skipLF := TRUE; END_IF;
            END_IF;
            IF NOT skipLF THEN
                IF count < 254 THEN
                    windows[window][count] := value;
                    count := count + 1;
                    windows[window][count] := 0;
                ELSE
                    Truncated := TRUE;
                END_IF;
            END_IF;
        END_IF;
    END_FOR;
END_FOR;
ByteArrayToString := windows[0];
ByteArrayToString_1 := windows[1];
ByteArrayToString_2 := windows[2];
ByteArrayToString_3 := windows[3];
ByteArrayToString_4 := windows[4];
ByteArrayToString_5 := windows[5];

END_FUNCTION

// ---- POUs/System/Functions/FC_TIAParseDINT.TcPOU
FUNCTION FC_TIAParseDINT : BOOL
VAR_INPUT
    Token : STRING(32);
END_VAR
VAR_OUTPUT
    Value : DINT;
END_VAR
VAR
    magnitude : LINT;
    negative : BOOL;
    cursor : INT;
    scan : INT;
    digit : INT;
    length : INT;
END_VAR

// Checked decimal conversion. Reject whitespace, fractions and overflow.
FC_TIAParseDINT := FALSE;
Value := 0;
magnitude := 0;
negative := FALSE;
cursor := 1;
length := LEN(Token);
IF length = 0 THEN RETURN; END_IF;
IF LEFT(Token, 1) = '-' THEN
    negative := TRUE;
    cursor := 2;
END_IF;
IF cursor > length THEN RETURN; END_IF;
IF (length - cursor + 1 > 1) AND (MID(Token, 1, cursor) = '0') THEN RETURN; END_IF;
FOR scan := cursor TO length DO
    digit := BYTE_TO_INT(Token[scan - 1]) - 48;
    IF (digit < 0) OR (digit > 9) THEN RETURN; END_IF;
    magnitude := magnitude * 10 + INT_TO_LINT(digit);
    // Early limit also bounds the next multiplication below LINT overflow.
    IF magnitude > LINT#2147483648 THEN RETURN; END_IF;
END_FOR;
IF negative THEN magnitude := -magnitude; END_IF;
IF magnitude > LINT#2147483647 THEN RETURN; END_IF;
Value := LINT_TO_DINT(magnitude);
FC_TIAParseDINT := TRUE;

END_FUNCTION

// ---- POUs/System/Functions/FC_TIAScalarToken.TcPOU
FUNCTION FC_TIAScalarToken : BOOL
VAR_INPUT
    FieldName : STRING(254);
    JsonStr : STRING(254);
END_VAR
VAR_OUTPUT
    Token : STRING(32);
END_VAR
VAR
    pattern : STRING(254);
    character : STRING(1);
    position : INT;
    cursor : INT;
    scan : INT;
    length : INT;
    valueStart : INT;
    previous : STRING(1);
END_VAR

// Restricted flat ASCII field extractor, not a general JSON parser.
// Require a complete scalar followed by ',' or '}'. Never accept truncation.
FC_TIAScalarToken := FALSE;
Token := '';
IF (LEN(FieldName) = 0) OR (LEN(FieldName) > 250) THEN RETURN; END_IF;
pattern := CONCAT(CONCAT('"', FieldName), '"');
position := FIND(JsonStr, pattern);
IF position = 0 THEN RETURN; END_IF;
// Reject field-name text inside a quoted value.
previous := '';
FOR scan := 1 TO position - 1 DO
    character := MID(JsonStr, 1, scan);
    IF (character <> ' ') AND (character <> '$T') AND
       (character <> '$R') AND (character <> '$N') THEN
        previous := character;
    END_IF;
END_FOR;
IF (previous <> '') AND (previous <> '{') AND (previous <> ',') THEN RETURN; END_IF;
length := LEN(JsonStr);
cursor := position + LEN(pattern);
FOR scan := cursor TO length DO
    character := MID(JsonStr, 1, scan);
    IF (character <> ' ') AND (character <> '$T') AND
       (character <> '$R') AND (character <> '$N') THEN EXIT; END_IF;
END_FOR;
IF scan > length THEN RETURN; END_IF;
IF MID(JsonStr, 1, scan) <> ':' THEN RETURN; END_IF;
cursor := scan + 1;
FOR scan := cursor TO length DO
    character := MID(JsonStr, 1, scan);
    IF (character <> ' ') AND (character <> '$T') AND
       (character <> '$R') AND (character <> '$N') THEN EXIT; END_IF;
END_FOR;
valueStart := scan;
FOR cursor := valueStart TO length DO
    character := MID(JsonStr, 1, cursor);
    IF (character = ',') OR (character = '}') THEN
        // Trim trailing JSON whitespace before extracting the token.
        position := cursor - 1;
        FOR scan := cursor - 1 TO valueStart BY -1 DO
            character := MID(JsonStr, 1, scan);
            IF (character <> ' ') AND (character <> '$T') AND
               (character <> '$R') AND (character <> '$N') THEN EXIT; END_IF;
            position := scan - 1;
        END_FOR;
        IF (position < valueStart) OR (position - valueStart + 1 > 32) THEN RETURN; END_IF;
        Token := MID(JsonStr, position - valueStart + 1, valueStart);
        FC_TIAScalarToken := TRUE;
        RETURN;
    END_IF;
END_FOR;

END_FUNCTION

// ---- POUs/System/Functions/FindBoolField.TcPOU
FUNCTION FindBoolField : BOOL
VAR_INPUT
    FieldName : STRING(254);
    JsonStr : STRING(254);
END_VAR
VAR_OUTPUT
    Valid : BOOL;
END_VAR
VAR
    token : STRING(32);
END_VAR

// Missing, malformed and false all return FALSE; inspect Valid to distinguish.
FindBoolField := FALSE;
Valid := FC_TIAScalarToken(FieldName := FieldName, JsonStr := JsonStr, Token => token);
IF NOT Valid THEN RETURN; END_IF;
Valid := (token = 'true') OR (token = 'false');
FindBoolField := token = 'true';

END_FUNCTION

// ---- POUs/System/Functions/FindDINTFieldFragmented.TcPOU
FUNCTION FindDINTFieldFragmented : DINT
VAR_INPUT
    FieldName : STRING(254);
    Str1 : STRING(254);
    Str2 : STRING(254);
END_VAR
VAR_OUTPUT
    Valid : BOOL;
END_VAR
VAR
    token : STRING(32);
    value : DINT;
    found : BOOL;
END_VAR

// Search complete fields in the reference's overlapping windows.
// Arbitrary concatenation of overlapping windows would corrupt payload data.
// A field split across both windows without a complete copy is rejected.
FindDINTFieldFragmented := -9999;
Valid := FALSE;
found := FC_TIAScalarToken(FieldName := FieldName, JsonStr := Str1, Token => token);
IF NOT found THEN
    found := FC_TIAScalarToken(FieldName := FieldName, JsonStr := Str2, Token => token);
END_IF;
IF NOT found THEN RETURN; END_IF;
Valid := FC_TIAParseDINT(Token := token, Value => value);
IF Valid THEN FindDINTFieldFragmented := value; END_IF;

END_FUNCTION

// ---- POUs/System/Functions/FindIntField.TcPOU
FUNCTION FindIntField : INT
VAR_INPUT
    FieldName : STRING(254);
    JsonStr : STRING(254);
END_VAR
VAR_OUTPUT
    Valid : BOOL;
END_VAR

FindIntField := FindINTFieldFragmented(FieldName := FieldName, Str1 := JsonStr, Str2 := '', Valid => Valid);

END_FUNCTION

